(* IEC 61131-3 sources: deprecated-refusr-repo/GP/Main/samples (part 5) *)

(* ---- 3-MUX_sappy-ovals-yanks.st ---- *)
(*
This code implements a shuffled multiplexer with 3 control bits.
The control bits are: Data[2], Data[4], Data[1]
The input bits are: Data[6], Data[3], Data[5], Data[7], Data[9], Data[8], Data[10], Data[11]

The symbolic expression is:
(((((((~((~(D[2]) & ~(D[4])) & ~(D[1])) | D[6]) & (~((D[2] & ~(D[4])) & ~(D[1])) | D[3])) & (~((~(D[2]) & D[4]) & ~(D[1])) | D[5])) & (~((D[2] & D[4]) & ~(D[1])) | D[7])) & (~((~(D[2]) & ~(D[4])) & D[1]) | D[9])) & (~((D[2] & ~(D[4])) & D[1]) | D[8])) & (~((~(D[2]) & D[4]) & D[1]) | D[10])) & (~((D[2] & D[4]) & D[1]) | D[11])

*)

FUNCTION_BLOCK F_CollectInput
  VAR_IN_OUT
      Data : ARRAY[1..15] OF BOOL;
  END_VAR
  VAR_INPUT
      TICK  : BOOL := 0;
      IN1   : BOOL := 0;
      IN2   : BOOL := 0;
      IN3   : BOOL := 0;
      IN4   : BOOL := 0;
      IN5   : BOOL := 0;
      RESET : BOOL := FALSE;
  END_VAR
  VAR_OUTPUT
      Finished : BOOL;
  END_VAR
  VAR
      j    : USINT := 1;
      tock : BOOL  := 0;
  END_VAR
  IF NOT RESET AND tock = NOT TICK THEN
      Data[j]   := IN1;
      Data[j+1] := IN2;
      Data[j+2] := IN3;
      Data[j+3] := IN4;
      Data[j+4] := IN5;
      j := j + 5;
      tock := TICK;
  ELSE
      j := 1;
      tock := 0;
  END_IF;
  Finished := (j > 15);
END_FUNCTION_BLOCK

PROGRAM Boiler
  VAR
    Data  : ARRAY[1..15] OF BOOL;
    Ready : BOOL;
    CollectInput : F_CollectInput;
  END_VAR
  VAR
    TICK     AT %IX1.0 : BOOL;
    IN1      AT %IX0.3 : BOOL;
    IN2      AT %IX0.4 : BOOL;
    IN3      AT %IX0.5 : BOOL;
    IN4      AT %IX0.6 : BOOL;
    IN5      AT %IX0.7 : BOOL;
    OutReady AT %QX0.0 : BOOL := FALSE;
    FeedNext AT %QX0.1 : BOOL := FALSE;
    Out      AT %QX0.2 : BOOL;
  END_VAR
  CollectInput(TICK:=TICK, IN1:=IN1, IN2:=IN2, IN3:=IN3, IN4:=IN4, IN5:=IN5);
  Ready := CollectInput.Finished;
  FeedNext := 1;
  IF Ready THEN
    Out := (((((((((NOT (((NOT D[2]) AND (NOT D[4])) AND (NOT D[1]))) OR D[6]) AND ((NOT ((D[2] AND (NOT D[4])) AND (NOT D[1]))) OR D[3])) AND ((NOT (((NOT D[2]) AND D[4]) AND (NOT D[1]))) OR D[5])) AND ((NOT ((D[2] AND D[4]) AND (NOT D[1]))) OR D[7])) AND ((NOT (((NOT D[2]) AND (NOT D[4])) AND D[1])) OR D[9])) AND ((NOT ((D[2] AND (NOT D[4])) AND D[1])) OR D[8])) AND ((NOT (((NOT D[2]) AND D[4]) AND D[1])) OR D[10])) AND ((NOT ((D[2] AND D[4]) AND D[1])) OR D[11]));
    OutReady := 1;
    CollectInput(RESET:=TRUE);
  END_IF;
END_PROGRAM

CONFIGURATION Config0
  RESOURCE Res0 ON PLC
    TASK task0(INTERVAL := T#20ms,PRIORITY := 0);
    PROGRAM instance0 WITH task0 : Boiler;
  END_RESOURCE
END_CONFIGURATION

(* ---- 3-MUX_scale-wants-nifty.st ---- *)
(*
This code implements a shuffled multiplexer with 3 control bits.
The control bits are: Data[2], Data[3], Data[5]
The input bits are: Data[1], Data[8], Data[9], Data[7], Data[4], Data[10], Data[6], Data[11]

The symbolic expression is:
(((((((~((~(D[2]) & ~(D[3])) & ~(D[5])) | D[1]) & (~((D[2] & ~(D[3])) & ~(D[5])) | D[8])) & (~((~(D[2]) & D[3]) & ~(D[5])) | D[9])) & (~((D[2] & D[3]) & ~(D[5])) | D[7])) & (~((~(D[2]) & ~(D[3])) & D[5]) | D[4])) & (~((D[2] & ~(D[3])) & D[5]) | D[10])) & (~((~(D[2]) & D[3]) & D[5]) | D[6])) & (~((D[2] & D[3]) & D[5]) | D[11])

*)

FUNCTION_BLOCK F_CollectInput
  VAR_IN_OUT
      Data : ARRAY[1..15] OF BOOL;
  END_VAR
  VAR_INPUT
      TICK  : BOOL := 0;
      IN1   : BOOL := 0;
      IN2   : BOOL := 0;
      IN3   : BOOL := 0;
      IN4   : BOOL := 0;
      IN5   : BOOL := 0;
      RESET : BOOL := FALSE;
  END_VAR
  VAR_OUTPUT
      Finished : BOOL;
  END_VAR
  VAR
      j    : USINT := 1;
      tock : BOOL  := 0;
  END_VAR
  IF NOT RESET AND tock = NOT TICK THEN
      Data[j]   := IN1;
      Data[j+1] := IN2;
      Data[j+2] := IN3;
      Data[j+3] := IN4;
      Data[j+4] := IN5;
      j := j + 5;
      tock := TICK;
  ELSE
      j := 1;
      tock := 0;
  END_IF;
  Finished := (j > 15);
END_FUNCTION_BLOCK

PROGRAM Boiler
  VAR
    Data  : ARRAY[1..15] OF BOOL;
    Ready : BOOL;
    CollectInput : F_CollectInput;
  END_VAR
  VAR
    TICK     AT %IX1.0 : BOOL;
    IN1      AT %IX0.3 : BOOL;
    IN2      AT %IX0.4 : BOOL;
    IN3      AT %IX0.5 : BOOL;
    IN4      AT %IX0.6 : BOOL;
    IN5      AT %IX0.7 : BOOL;
    OutReady AT %QX0.0 : BOOL := FALSE;
    FeedNext AT %QX0.1 : BOOL := FALSE;
    Out      AT %QX0.2 : BOOL;
  END_VAR
  CollectInput(TICK:=TICK, IN1:=IN1, IN2:=IN2, IN3:=IN3, IN4:=IN4, IN5:=IN5);
  Ready := CollectInput.Finished;
  FeedNext := 1;
  IF Ready THEN
    Out := (((((((((NOT (((NOT D[2]) AND (NOT D[3])) AND (NOT D[5]))) OR D[1]) AND ((NOT ((D[2] AND (NOT D[3])) AND (NOT D[5]))) OR D[8])) AND ((NOT (((NOT D[2]) AND D[3]) AND (NOT D[5]))) OR D[9])) AND ((NOT ((D[2] AND D[3]) AND (NOT D[5]))) OR D[7])) AND ((NOT (((NOT D[2]) AND (NOT D[3])) AND D[5])) OR D[4])) AND ((NOT ((D[2] AND (NOT D[3])) AND D[5])) OR D[10])) AND ((NOT (((NOT D[2]) AND D[3]) AND D[5])) OR D[6])) AND ((NOT ((D[2] AND D[3]) AND D[5])) OR D[11]));
    OutReady := 1;
    CollectInput(RESET:=TRUE);
  END_IF;
END_PROGRAM

CONFIGURATION Config0
  RESOURCE Res0 ON PLC
    TASK task0(INTERVAL := T#20ms,PRIORITY := 0);
    PROGRAM instance0 WITH task0 : Boiler;
  END_RESOURCE
END_CONFIGURATION

(* ---- 3-MUX_scion-boxer-krona.st ---- *)
(*
This code implements a shuffled multiplexer with 3 control bits.
The control bits are: Data[3], Data[5], Data[4]
The input bits are: Data[1], Data[2], Data[9], Data[6], Data[10], Data[7], Data[11], Data[8]

The symbolic expression is:
(((((((~((~(D[3]) & ~(D[5])) & ~(D[4])) | D[1]) & (~((D[3] & ~(D[5])) & ~(D[4])) | D[2])) & (~((~(D[3]) & D[5]) & ~(D[4])) | D[9])) & (~((D[3] & D[5]) & ~(D[4])) | D[6])) & (~((~(D[3]) & ~(D[5])) & D[4]) | D[10])) & (~((D[3] & ~(D[5])) & D[4]) | D[7])) & (~((~(D[3]) & D[5]) & D[4]) | D[11])) & (~((D[3] & D[5]) & D[4]) | D[8])

*)

FUNCTION_BLOCK F_CollectInput
  VAR_IN_OUT
      Data : ARRAY[1..15] OF BOOL;
  END_VAR
  VAR_INPUT
      TICK  : BOOL := 0;
      IN1   : BOOL := 0;
      IN2   : BOOL := 0;
      IN3   : BOOL := 0;
      IN4   : BOOL := 0;
      IN5   : BOOL := 0;
      RESET : BOOL := FALSE;
  END_VAR
  VAR_OUTPUT
      Finished : BOOL;
  END_VAR
  VAR
      j    : USINT := 1;
      tock : BOOL  := 0;
  END_VAR
  IF NOT RESET AND tock = NOT TICK THEN
      Data[j]   := IN1;
      Data[j+1] := IN2;
      Data[j+2] := IN3;
      Data[j+3] := IN4;
      Data[j+4] := IN5;
      j := j + 5;
      tock := TICK;
  ELSE
      j := 1;
      tock := 0;
  END_IF;
  Finished := (j > 15);
END_FUNCTION_BLOCK

PROGRAM Boiler
  VAR
    Data  : ARRAY[1..15] OF BOOL;
    Ready : BOOL;
    CollectInput : F_CollectInput;
  END_VAR
  VAR
    TICK     AT %IX1.0 : BOOL;
    IN1      AT %IX0.3 : BOOL;
    IN2      AT %IX0.4 : BOOL;
    IN3      AT %IX0.5 : BOOL;
    IN4      AT %IX0.6 : BOOL;
    IN5      AT %IX0.7 : BOOL;
    OutReady AT %QX0.0 : BOOL := FALSE;
    FeedNext AT %QX0.1 : BOOL := FALSE;
    Out      AT %QX0.2 : BOOL;
  END_VAR
  CollectInput(TICK:=TICK, IN1:=IN1, IN2:=IN2, IN3:=IN3, IN4:=IN4, IN5:=IN5);
  Ready := CollectInput.Finished;
  FeedNext := 1;
  IF Ready THEN
    Out := (((((((((NOT (((NOT D[3]) AND (NOT D[5])) AND (NOT D[4]))) OR D[1]) AND ((NOT ((D[3] AND (NOT D[5])) AND (NOT D[4]))) OR D[2])) AND ((NOT (((NOT D[3]) AND D[5]) AND (NOT D[4]))) OR D[9])) AND ((NOT ((D[3] AND D[5]) AND (NOT D[4]))) OR D[6])) AND ((NOT (((NOT D[3]) AND (NOT D[5])) AND D[4])) OR D[10])) AND ((NOT ((D[3] AND (NOT D[5])) AND D[4])) OR D[7])) AND ((NOT (((NOT D[3]) AND D[5]) AND D[4])) OR D[11])) AND ((NOT ((D[3] AND D[5]) AND D[4])) OR D[8]));
    OutReady := 1;
    CollectInput(RESET:=TRUE);
  END_IF;
END_PROGRAM

CONFIGURATION Config0
  RESOURCE Res0 ON PLC
    TASK task0(INTERVAL := T#20ms,PRIORITY := 0);
    PROGRAM instance0 WITH task0 : Boiler;
  END_RESOURCE
END_CONFIGURATION

(* ---- 3-MUX_sects-chimp-tilth.st ---- *)
(*
This code implements a shuffled multiplexer with 3 control bits.
The control bits are: Data[2], Data[1], Data[5]
The input bits are: Data[3], Data[4], Data[6], Data[9], Data[7], Data[10], Data[11], Data[8]

The symbolic expression is:
(((((((~((~(D[2]) & ~(D[1])) & ~(D[5])) | D[3]) & (~((D[2] & ~(D[1])) & ~(D[5])) | D[4])) & (~((~(D[2]) & D[1]) & ~(D[5])) | D[6])) & (~((D[2] & D[1]) & ~(D[5])) | D[9])) & (~((~(D[2]) & ~(D[1])) & D[5]) | D[7])) & (~((D[2] & ~(D[1])) & D[5]) | D[10])) & (~((~(D[2]) & D[1]) & D[5]) | D[11])) & (~((D[2] & D[1]) & D[5]) | D[8])

*)

FUNCTION_BLOCK F_CollectInput
  VAR_IN_OUT
      Data : ARRAY[1..15] OF BOOL;
  END_VAR
  VAR_INPUT
      TICK  : BOOL := 0;
      IN1   : BOOL := 0;
      IN2   : BOOL := 0;
      IN3   : BOOL := 0;
      IN4   : BOOL := 0;
      IN5   : BOOL := 0;
      RESET : BOOL := FALSE;
  END_VAR
  VAR_OUTPUT
      Finished : BOOL;
  END_VAR
  VAR
      j    : USINT := 1;
      tock : BOOL  := 0;
  END_VAR
  IF NOT RESET AND tock = NOT TICK THEN
      Data[j]   := IN1;
      Data[j+1] := IN2;
      Data[j+2] := IN3;
      Data[j+3] := IN4;
      Data[j+4] := IN5;
      j := j + 5;
      tock := TICK;
  ELSE
      j := 1;
      tock := 0;
  END_IF;
  Finished := (j > 15);
END_FUNCTION_BLOCK

PROGRAM Boiler
  VAR
    Data  : ARRAY[1..15] OF BOOL;
    Ready : BOOL;
    CollectInput : F_CollectInput;
  END_VAR
  VAR
    TICK     AT %IX1.0 : BOOL;
    IN1      AT %IX0.3 : BOOL;
    IN2      AT %IX0.4 : BOOL;
    IN3      AT %IX0.5 : BOOL;
    IN4      AT %IX0.6 : BOOL;
    IN5      AT %IX0.7 : BOOL;
    OutReady AT %QX0.0 : BOOL := FALSE;
    FeedNext AT %QX0.1 : BOOL := FALSE;
    Out      AT %QX0.2 : BOOL;
  END_VAR
  CollectInput(TICK:=TICK, IN1:=IN1, IN2:=IN2, IN3:=IN3, IN4:=IN4, IN5:=IN5);
  Ready := CollectInput.Finished;
  FeedNext := 1;
  IF Ready THEN
    Out := (((((((((NOT (((NOT D[2]) AND (NOT D[1])) AND (NOT D[5]))) OR D[3]) AND ((NOT ((D[2] AND (NOT D[1])) AND (NOT D[5]))) OR D[4])) AND ((NOT (((NOT D[2]) AND D[1]) AND (NOT D[5]))) OR D[6])) AND ((NOT ((D[2] AND D[1]) AND (NOT D[5]))) OR D[9])) AND ((NOT (((NOT D[2]) AND (NOT D[1])) AND D[5])) OR D[7])) AND ((NOT ((D[2] AND (NOT D[1])) AND D[5])) OR D[10])) AND ((NOT (((NOT D[2]) AND D[1]) AND D[5])) OR D[11])) AND ((NOT ((D[2] AND D[1]) AND D[5])) OR D[8]));
    OutReady := 1;
    CollectInput(RESET:=TRUE);
  END_IF;
END_PROGRAM

CONFIGURATION Config0
  RESOURCE Res0 ON PLC
    TASK task0(INTERVAL := T#20ms,PRIORITY := 0);
    PROGRAM instance0 WITH task0 : Boiler;
  END_RESOURCE
END_CONFIGURATION

(* ---- 3-MUX_seems-zebra-casus.st ---- *)
(*
This code implements a shuffled multiplexer with 3 control bits.
The control bits are: Data[1], Data[2], Data[3]
The input bits are: Data[7], Data[5], Data[4], Data[6], Data[8], Data[9], Data[10], Data[11]

The symbolic expression is:
(((((((~((~(D[1]) & ~(D[2])) & ~(D[3])) | D[7]) & (~((D[1] & ~(D[2])) & ~(D[3])) | D[5])) & (~((~(D[1]) & D[2]) & ~(D[3])) | D[4])) & (~((D[1] & D[2]) & ~(D[3])) | D[6])) & (~((~(D[1]) & ~(D[2])) & D[3]) | D[8])) & (~((D[1] & ~(D[2])) & D[3]) | D[9])) & (~((~(D[1]) & D[2]) & D[3]) | D[10])) & (~((D[1] & D[2]) & D[3]) | D[11])

*)

FUNCTION_BLOCK F_CollectInput
  VAR_IN_OUT
      Data : ARRAY[1..15] OF BOOL;
  END_VAR
  VAR_INPUT
      TICK  : BOOL := 0;
      IN1   : BOOL := 0;
      IN2   : BOOL := 0;
      IN3   : BOOL := 0;
      IN4   : BOOL := 0;
      IN5   : BOOL := 0;
      RESET : BOOL := FALSE;
  END_VAR
  VAR_OUTPUT
      Finished : BOOL;
  END_VAR
  VAR
      j    : USINT := 1;
      tock : BOOL  := 0;
  END_VAR
  IF NOT RESET AND tock = NOT TICK THEN
      Data[j]   := IN1;
      Data[j+1] := IN2;
      Data[j+2] := IN3;
      Data[j+3] := IN4;
      Data[j+4] := IN5;
      j := j + 5;
      tock := TICK;
  ELSE
      j := 1;
      tock := 0;
  END_IF;
  Finished := (j > 15);
END_FUNCTION_BLOCK

PROGRAM Boiler
  VAR
    Data  : ARRAY[1..15] OF BOOL;
    Ready : BOOL;
    CollectInput : F_CollectInput;
  END_VAR
  VAR
    TICK     AT %IX1.0 : BOOL;
    IN1      AT %IX0.3 : BOOL;
    IN2      AT %IX0.4 : BOOL;
    IN3      AT %IX0.5 : BOOL;
    IN4      AT %IX0.6 : BOOL;
    IN5      AT %IX0.7 : BOOL;
    OutReady AT %QX0.0 : BOOL := FALSE;
    FeedNext AT %QX0.1 : BOOL := FALSE;
    Out      AT %QX0.2 : BOOL;
  END_VAR
  CollectInput(TICK:=TICK, IN1:=IN1, IN2:=IN2, IN3:=IN3, IN4:=IN4, IN5:=IN5);
  Ready := CollectInput.Finished;
  FeedNext := 1;
  IF Ready THEN
    Out := (((((((((NOT (((NOT D[1]) AND (NOT D[2])) AND (NOT D[3]))) OR D[7]) AND ((NOT ((D[1] AND (NOT D[2])) AND (NOT D[3]))) OR D[5])) AND ((NOT (((NOT D[1]) AND D[2]) AND (NOT D[3]))) OR D[4])) AND ((NOT ((D[1] AND D[2]) AND (NOT D[3]))) OR D[6])) AND ((NOT (((NOT D[1]) AND (NOT D[2])) AND D[3])) OR D[8])) AND ((NOT ((D[1] AND (NOT D[2])) AND D[3])) OR D[9])) AND ((NOT (((NOT D[1]) AND D[2]) AND D[3])) OR D[10])) AND ((NOT ((D[1] AND D[2]) AND D[3])) OR D[11]));
    OutReady := 1;
    CollectInput(RESET:=TRUE);
  END_IF;
END_PROGRAM

CONFIGURATION Config0
  RESOURCE Res0 ON PLC
    TASK task0(INTERVAL := T#20ms,PRIORITY := 0);
    PROGRAM instance0 WITH task0 : Boiler;
  END_RESOURCE
END_CONFIGURATION

(* ---- 3-MUX_shunt-caret-reedy.st ---- *)
(*
This code implements a shuffled multiplexer with 3 control bits.
The control bits are: Data[5], Data[3], Data[1]
The input bits are: Data[4], Data[6], Data[8], Data[7], Data[10], Data[11], Data[9], Data[2]

The symbolic expression is:
(((((((~((~(D[5]) & ~(D[3])) & ~(D[1])) | D[4]) & (~((D[5] & ~(D[3])) & ~(D[1])) | D[6])) & (~((~(D[5]) & D[3]) & ~(D[1])) | D[8])) & (~((D[5] & D[3]) & ~(D[1])) | D[7])) & (~((~(D[5]) & ~(D[3])) & D[1]) | D[10])) & (~((D[5] & ~(D[3])) & D[1]) | D[11])) & (~((~(D[5]) & D[3]) & D[1]) | D[9])) & (~((D[5] & D[3]) & D[1]) | D[2])

*)

FUNCTION_BLOCK F_CollectInput
  VAR_IN_OUT
      Data : ARRAY[1..15] OF BOOL;
  END_VAR
  VAR_INPUT
      TICK  : BOOL := 0;
      IN1   : BOOL := 0;
      IN2   : BOOL := 0;
      IN3   : BOOL := 0;
      IN4   : BOOL := 0;
      IN5   : BOOL := 0;
      RESET : BOOL := FALSE;
  END_VAR
  VAR_OUTPUT
      Finished : BOOL;
  END_VAR
  VAR
      j    : USINT := 1;
      tock : BOOL  := 0;
  END_VAR
  IF NOT RESET AND tock = NOT TICK THEN
      Data[j]   := IN1;
      Data[j+1] := IN2;
      Data[j+2] := IN3;
      Data[j+3] := IN4;
      Data[j+4] := IN5;
      j := j + 5;
      tock := TICK;
  ELSE
      j := 1;
      tock := 0;
  END_IF;
  Finished := (j > 15);
END_FUNCTION_BLOCK

PROGRAM Boiler
  VAR
    Data  : ARRAY[1..15] OF BOOL;
    Ready : BOOL;
    CollectInput : F_CollectInput;
  END_VAR
  VAR
    TICK     AT %IX1.0 : BOOL;
    IN1      AT %IX0.3 : BOOL;
    IN2      AT %IX0.4 : BOOL;
    IN3      AT %IX0.5 : BOOL;
    IN4      AT %IX0.6 : BOOL;
    IN5      AT %IX0.7 : BOOL;
    OutReady AT %QX0.0 : BOOL := FALSE;
    FeedNext AT %QX0.1 : BOOL := FALSE;
    Out      AT %QX0.2 : BOOL;
  END_VAR
  CollectInput(TICK:=TICK, IN1:=IN1, IN2:=IN2, IN3:=IN3, IN4:=IN4, IN5:=IN5);
  Ready := CollectInput.Finished;
  FeedNext := 1;
  IF Ready THEN
    Out := (((((((((NOT (((NOT D[5]) AND (NOT D[3])) AND (NOT D[1]))) OR D[4]) AND ((NOT ((D[5] AND (NOT D[3])) AND (NOT D[1]))) OR D[6])) AND ((NOT (((NOT D[5]) AND D[3]) AND (NOT D[1]))) OR D[8])) AND ((NOT ((D[5] AND D[3]) AND (NOT D[1]))) OR D[7])) AND ((NOT (((NOT D[5]) AND (NOT D[3])) AND D[1])) OR D[10])) AND ((NOT ((D[5] AND (NOT D[3])) AND D[1])) OR D[11])) AND ((NOT (((NOT D[5]) AND D[3]) AND D[1])) OR D[9])) AND ((NOT ((D[5] AND D[3]) AND D[1])) OR D[2]));
    OutReady := 1;
    CollectInput(RESET:=TRUE);
  END_IF;
END_PROGRAM

CONFIGURATION Config0
  RESOURCE Res0 ON PLC
    TASK task0(INTERVAL := T#20ms,PRIORITY := 0);
    PROGRAM instance0 WITH task0 : Boiler;
  END_RESOURCE
END_CONFIGURATION

(* ---- 3-MUX_slums-noted-letup.st ---- *)
(*
This code implements a shuffled multiplexer with 3 control bits.
The control bits are: Data[3], Data[4], Data[1]
The input bits are: Data[9], Data[2], Data[11], Data[5], Data[7], Data[8], Data[6], Data[10]

The symbolic expression is:
(((((((~((~(D[3]) & ~(D[4])) & ~(D[1])) | D[9]) & (~((D[3] & ~(D[4])) & ~(D[1])) | D[2])) & (~((~(D[3]) & D[4]) & ~(D[1])) | D[11])) & (~((D[3] & D[4]) & ~(D[1])) | D[5])) & (~((~(D[3]) & ~(D[4])) & D[1]) | D[7])) & (~((D[3] & ~(D[4])) & D[1]) | D[8])) & (~((~(D[3]) & D[4]) & D[1]) | D[6])) & (~((D[3] & D[4]) & D[1]) | D[10])

*)

FUNCTION_BLOCK F_CollectInput
  VAR_IN_OUT
      Data : ARRAY[1..15] OF BOOL;
  END_VAR
  VAR_INPUT
      TICK  : BOOL := 0;
      IN1   : BOOL := 0;
      IN2   : BOOL := 0;
      IN3   : BOOL := 0;
      IN4   : BOOL := 0;
      IN5   : BOOL := 0;
      RESET : BOOL := FALSE;
  END_VAR
  VAR_OUTPUT
      Finished : BOOL;
  END_VAR
  VAR
      j    : USINT := 1;
      tock : BOOL  := 0;
  END_VAR
  IF NOT RESET AND tock = NOT TICK THEN
      Data[j]   := IN1;
      Data[j+1] := IN2;
      Data[j+2] := IN3;
      Data[j+3] := IN4;
      Data[j+4] := IN5;
      j := j + 5;
      tock := TICK;
  ELSE
      j := 1;
      tock := 0;
  END_IF;
  Finished := (j > 15);
END_FUNCTION_BLOCK

PROGRAM Boiler
  VAR
    Data  : ARRAY[1..15] OF BOOL;
    Ready : BOOL;
    CollectInput : F_CollectInput;
  END_VAR
  VAR
    TICK     AT %IX1.0 : BOOL;
    IN1      AT %IX0.3 : BOOL;
    IN2      AT %IX0.4 : BOOL;
    IN3      AT %IX0.5 : BOOL;
    IN4      AT %IX0.6 : BOOL;
    IN5      AT %IX0.7 : BOOL;
    OutReady AT %QX0.0 : BOOL := FALSE;
    FeedNext AT %QX0.1 : BOOL := FALSE;
    Out      AT %QX0.2 : BOOL;
  END_VAR
  CollectInput(TICK:=TICK, IN1:=IN1, IN2:=IN2, IN3:=IN3, IN4:=IN4, IN5:=IN5);
  Ready := CollectInput.Finished;
  FeedNext := 1;
  IF Ready THEN
    Out := (((((((((NOT (((NOT D[3]) AND (NOT D[4])) AND (NOT D[1]))) OR D[9]) AND ((NOT ((D[3] AND (NOT D[4])) AND (NOT D[1]))) OR D[2])) AND ((NOT (((NOT D[3]) AND D[4]) AND (NOT D[1]))) OR D[11])) AND ((NOT ((D[3] AND D[4]) AND (NOT D[1]))) OR D[5])) AND ((NOT (((NOT D[3]) AND (NOT D[4])) AND D[1])) OR D[7])) AND ((NOT ((D[3] AND (NOT D[4])) AND D[1])) OR D[8])) AND ((NOT (((NOT D[3]) AND D[4]) AND D[1])) OR D[6])) AND ((NOT ((D[3] AND D[4]) AND D[1])) OR D[10]));
    OutReady := 1;
    CollectInput(RESET:=TRUE);
  END_IF;
END_PROGRAM

CONFIGURATION Config0
  RESOURCE Res0 ON PLC
    TASK task0(INTERVAL := T#20ms,PRIORITY := 0);
    PROGRAM instance0 WITH task0 : Boiler;
  END_RESOURCE
END_CONFIGURATION

(* ---- 3-MUX_sonny-vised-eying.st ---- *)
(*
This code implements a shuffled multiplexer with 3 control bits.
The control bits are: Data[2], Data[1], Data[4]
The input bits are: Data[3], Data[7], Data[6], Data[8], Data[5], Data[9], Data[11], Data[10]

The symbolic expression is:
(((((((~((~(D[2]) & ~(D[1])) & ~(D[4])) | D[3]) & (~((D[2] & ~(D[1])) & ~(D[4])) | D[7])) & (~((~(D[2]) & D[1]) & ~(D[4])) | D[6])) & (~((D[2] & D[1]) & ~(D[4])) | D[8])) & (~((~(D[2]) & ~(D[1])) & D[4]) | D[5])) & (~((D[2] & ~(D[1])) & D[4]) | D[9])) & (~((~(D[2]) & D[1]) & D[4]) | D[11])) & (~((D[2] & D[1]) & D[4]) | D[10])

*)

FUNCTION_BLOCK F_CollectInput
  VAR_IN_OUT
      Data : ARRAY[1..15] OF BOOL;
  END_VAR
  VAR_INPUT
      TICK  : BOOL := 0;
      IN1   : BOOL := 0;
      IN2   : BOOL := 0;
      IN3   : BOOL := 0;
      IN4   : BOOL := 0;
      IN5   : BOOL := 0;
      RESET : BOOL := FALSE;
  END_VAR
  VAR_OUTPUT
      Finished : BOOL;
  END_VAR
  VAR
      j    : USINT := 1;
      tock : BOOL  := 0;
  END_VAR
  IF NOT RESET AND tock = NOT TICK THEN
      Data[j]   := IN1;
      Data[j+1] := IN2;
      Data[j+2] := IN3;
      Data[j+3] := IN4;
      Data[j+4] := IN5;
      j := j + 5;
      tock := TICK;
  ELSE
      j := 1;
      tock := 0;
  END_IF;
  Finished := (j > 15);
END_FUNCTION_BLOCK

PROGRAM Boiler
  VAR
    Data  : ARRAY[1..15] OF BOOL;
    Ready : BOOL;
    CollectInput : F_CollectInput;
  END_VAR
  VAR
    TICK     AT %IX1.0 : BOOL;
    IN1      AT %IX0.3 : BOOL;
    IN2      AT %IX0.4 : BOOL;
    IN3      AT %IX0.5 : BOOL;
    IN4      AT %IX0.6 : BOOL;
    IN5      AT %IX0.7 : BOOL;
    OutReady AT %QX0.0 : BOOL := FALSE;
    FeedNext AT %QX0.1 : BOOL := FALSE;
    Out      AT %QX0.2 : BOOL;
  END_VAR
  CollectInput(TICK:=TICK, IN1:=IN1, IN2:=IN2, IN3:=IN3, IN4:=IN4, IN5:=IN5);
  Ready := CollectInput.Finished;
  FeedNext := 1;
  IF Ready THEN
    Out := (((((((((NOT (((NOT D[2]) AND (NOT D[1])) AND (NOT D[4]))) OR D[3]) AND ((NOT ((D[2] AND (NOT D[1])) AND (NOT D[4]))) OR D[7])) AND ((NOT (((NOT D[2]) AND D[1]) AND (NOT D[4]))) OR D[6])) AND ((NOT ((D[2] AND D[1]) AND (NOT D[4]))) OR D[8])) AND ((NOT (((NOT D[2]) AND (NOT D[1])) AND D[4])) OR D[5])) AND ((NOT ((D[2] AND (NOT D[1])) AND D[4])) OR D[9])) AND ((NOT (((NOT D[2]) AND D[1]) AND D[4])) OR D[11])) AND ((NOT ((D[2] AND D[1]) AND D[4])) OR D[10]));
    OutReady := 1;
    CollectInput(RESET:=TRUE);
  END_IF;
END_PROGRAM

CONFIGURATION Config0
  RESOURCE Res0 ON PLC
    TASK task0(INTERVAL := T#20ms,PRIORITY := 0);
    PROGRAM instance0 WITH task0 : Boiler;
  END_RESOURCE
END_CONFIGURATION

(* ---- 3-MUX_spark-lithe-swans.st ---- *)
(*
This code implements a shuffled multiplexer with 3 control bits.
The control bits are: Data[4], Data[3], Data[1]
The input bits are: Data[5], Data[6], Data[2], Data[7], Data[10], Data[8], Data[9], Data[11]

The symbolic expression is:
(((((((~((~(D[4]) & ~(D[3])) & ~(D[1])) | D[5]) & (~((D[4] & ~(D[3])) & ~(D[1])) | D[6])) & (~((~(D[4]) & D[3]) & ~(D[1])) | D[2])) & (~((D[4] & D[3]) & ~(D[1])) | D[7])) & (~((~(D[4]) & ~(D[3])) & D[1]) | D[10])) & (~((D[4] & ~(D[3])) & D[1]) | D[8])) & (~((~(D[4]) & D[3]) & D[1]) | D[9])) & (~((D[4] & D[3]) & D[1]) | D[11])

*)

FUNCTION_BLOCK F_CollectInput
  VAR_IN_OUT
      Data : ARRAY[1..15] OF BOOL;
  END_VAR
  VAR_INPUT
      TICK  : BOOL := 0;
      IN1   : BOOL := 0;
      IN2   : BOOL := 0;
      IN3   : BOOL := 0;
      IN4   : BOOL := 0;
      IN5   : BOOL := 0;
      RESET : BOOL := FALSE;
  END_VAR
  VAR_OUTPUT
      Finished : BOOL;
  END_VAR
  VAR
      j    : USINT := 1;
      tock : BOOL  := 0;
  END_VAR
  IF NOT RESET AND tock = NOT TICK THEN
      Data[j]   := IN1;
      Data[j+1] := IN2;
      Data[j+2] := IN3;
      Data[j+3] := IN4;
      Data[j+4] := IN5;
      j := j + 5;
      tock := TICK;
  ELSE
      j := 1;
      tock := 0;
  END_IF;
  Finished := (j > 15);
END_FUNCTION_BLOCK

PROGRAM Boiler
  VAR
    Data  : ARRAY[1..15] OF BOOL;
    Ready : BOOL;
    CollectInput : F_CollectInput;
  END_VAR
  VAR
    TICK     AT %IX1.0 : BOOL;
    IN1      AT %IX0.3 : BOOL;
    IN2      AT %IX0.4 : BOOL;
    IN3      AT %IX0.5 : BOOL;
    IN4      AT %IX0.6 : BOOL;
    IN5      AT %IX0.7 : BOOL;
    OutReady AT %QX0.0 : BOOL := FALSE;
    FeedNext AT %QX0.1 : BOOL := FALSE;
    Out      AT %QX0.2 : BOOL;
  END_VAR
  CollectInput(TICK:=TICK, IN1:=IN1, IN2:=IN2, IN3:=IN3, IN4:=IN4, IN5:=IN5);
  Ready := CollectInput.Finished;
  FeedNext := 1;
  IF Ready THEN
    Out := (((((((((NOT (((NOT D[4]) AND (NOT D[3])) AND (NOT D[1]))) OR D[5]) AND ((NOT ((D[4] AND (NOT D[3])) AND (NOT D[1]))) OR D[6])) AND ((NOT (((NOT D[4]) AND D[3]) AND (NOT D[1]))) OR D[2])) AND ((NOT ((D[4] AND D[3]) AND (NOT D[1]))) OR D[7])) AND ((NOT (((NOT D[4]) AND (NOT D[3])) AND D[1])) OR D[10])) AND ((NOT ((D[4] AND (NOT D[3])) AND D[1])) OR D[8])) AND ((NOT (((NOT D[4]) AND D[3]) AND D[1])) OR D[9])) AND ((NOT ((D[4] AND D[3]) AND D[1])) OR D[11]));
    OutReady := 1;
    CollectInput(RESET:=TRUE);
  END_IF;
END_PROGRAM

CONFIGURATION Config0
  RESOURCE Res0 ON PLC
    TASK task0(INTERVAL := T#20ms,PRIORITY := 0);
    PROGRAM instance0 WITH task0 : Boiler;
  END_RESOURCE
END_CONFIGURATION

(* ---- 3-MUX_spoof-lawns-sylph.st ---- *)
(*
This code implements a shuffled multiplexer with 3 control bits.
The control bits are: Data[2], Data[1], Data[3]
The input bits are: Data[4], Data[7], Data[8], Data[5], Data[9], Data[6], Data[10], Data[11]

The symbolic expression is:
(((((((~((~(D[2]) & ~(D[1])) & ~(D[3])) | D[4]) & (~((D[2] & ~(D[1])) & ~(D[3])) | D[7])) & (~((~(D[2]) & D[1]) & ~(D[3])) | D[8])) & (~((D[2] & D[1]) & ~(D[3])) | D[5])) & (~((~(D[2]) & ~(D[1])) & D[3]) | D[9])) & (~((D[2] & ~(D[1])) & D[3]) | D[6])) & (~((~(D[2]) & D[1]) & D[3]) | D[10])) & (~((D[2] & D[1]) & D[3]) | D[11])

*)

FUNCTION_BLOCK F_CollectInput
  VAR_IN_OUT
      Data : ARRAY[1..15] OF BOOL;
  END_VAR
  VAR_INPUT
      TICK  : BOOL := 0;
      IN1   : BOOL := 0;
      IN2   : BOOL := 0;
      IN3   : BOOL := 0;
      IN4   : BOOL := 0;
      IN5   : BOOL := 0;
      RESET : BOOL := FALSE;
  END_VAR
  VAR_OUTPUT
      Finished : BOOL;
  END_VAR
  VAR
      j    : USINT := 1;
      tock : BOOL  := 0;
  END_VAR
  IF NOT RESET AND tock = NOT TICK THEN
      Data[j]   := IN1;
      Data[j+1] := IN2;
      Data[j+2] := IN3;
      Data[j+3] := IN4;
      Data[j+4] := IN5;
      j := j + 5;
      tock := TICK;
  ELSE
      j := 1;
      tock := 0;
  END_IF;
  Finished := (j > 15);
END_FUNCTION_BLOCK

PROGRAM Boiler
  VAR
    Data  : ARRAY[1..15] OF BOOL;
    Ready : BOOL;
    CollectInput : F_CollectInput;
  END_VAR
  VAR
    TICK     AT %IX1.0 : BOOL;
    IN1      AT %IX0.3 : BOOL;
    IN2      AT %IX0.4 : BOOL;
    IN3      AT %IX0.5 : BOOL;
    IN4      AT %IX0.6 : BOOL;
    IN5      AT %IX0.7 : BOOL;
    OutReady AT %QX0.0 : BOOL := FALSE;
    FeedNext AT %QX0.1 : BOOL := FALSE;
    Out      AT %QX0.2 : BOOL;
  END_VAR
  CollectInput(TICK:=TICK, IN1:=IN1, IN2:=IN2, IN3:=IN3, IN4:=IN4, IN5:=IN5);
  Ready := CollectInput.Finished;
  FeedNext := 1;
  IF Ready THEN
    Out := (((((((((NOT (((NOT D[2]) AND (NOT D[1])) AND (NOT D[3]))) OR D[4]) AND ((NOT ((D[2] AND (NOT D[1])) AND (NOT D[3]))) OR D[7])) AND ((NOT (((NOT D[2]) AND D[1]) AND (NOT D[3]))) OR D[8])) AND ((NOT ((D[2] AND D[1]) AND (NOT D[3]))) OR D[5])) AND ((NOT (((NOT D[2]) AND (NOT D[1])) AND D[3])) OR D[9])) AND ((NOT ((D[2] AND (NOT D[1])) AND D[3])) OR D[6])) AND ((NOT (((NOT D[2]) AND D[1]) AND D[3])) OR D[10])) AND ((NOT ((D[2] AND D[1]) AND D[3])) OR D[11]));
    OutReady := 1;
    CollectInput(RESET:=TRUE);
  END_IF;
END_PROGRAM

CONFIGURATION Config0
  RESOURCE Res0 ON PLC
    TASK task0(INTERVAL := T#20ms,PRIORITY := 0);
    PROGRAM instance0 WITH task0 : Boiler;
  END_RESOURCE
END_CONFIGURATION

(* ---- 3-MUX_steer-patsy-bored.st ---- *)
(*
This code implements a shuffled multiplexer with 3 control bits.
The control bits are: Data[3], Data[1], Data[2]
The input bits are: Data[5], Data[4], Data[6], Data[9], Data[7], Data[11], Data[8], Data[10]

The symbolic expression is:
(((((((~((~(D[3]) & ~(D[1])) & ~(D[2])) | D[5]) & (~((D[3] & ~(D[1])) & ~(D[2])) | D[4])) & (~((~(D[3]) & D[1]) & ~(D[2])) | D[6])) & (~((D[3] & D[1]) & ~(D[2])) | D[9])) & (~((~(D[3]) & ~(D[1])) & D[2]) | D[7])) & (~((D[3] & ~(D[1])) & D[2]) | D[11])) & (~((~(D[3]) & D[1]) & D[2]) | D[8])) & (~((D[3] & D[1]) & D[2]) | D[10])

*)

FUNCTION_BLOCK F_CollectInput
  VAR_IN_OUT
      Data : ARRAY[1..15] OF BOOL;
  END_VAR
  VAR_INPUT
      TICK  : BOOL := 0;
      IN1   : BOOL := 0;
      IN2   : BOOL := 0;
      IN3   : BOOL := 0;
      IN4   : BOOL := 0;
      IN5   : BOOL := 0;
      RESET : BOOL := FALSE;
  END_VAR
  VAR_OUTPUT
      Finished : BOOL;
  END_VAR
  VAR
      j    : USINT := 1;
      tock : BOOL  := 0;
  END_VAR
  IF NOT RESET AND tock = NOT TICK THEN
      Data[j]   := IN1;
      Data[j+1] := IN2;
      Data[j+2] := IN3;
      Data[j+3] := IN4;
      Data[j+4] := IN5;
      j := j + 5;
      tock := TICK;
  ELSE
      j := 1;
      tock := 0;
  END_IF;
  Finished := (j > 15);
END_FUNCTION_BLOCK

PROGRAM Boiler
  VAR
    Data  : ARRAY[1..15] OF BOOL;
    Ready : BOOL;
    CollectInput : F_CollectInput;
  END_VAR
  VAR
    TICK     AT %IX1.0 : BOOL;
    IN1      AT %IX0.3 : BOOL;
    IN2      AT %IX0.4 : BOOL;
    IN3      AT %IX0.5 : BOOL;
    IN4      AT %IX0.6 : BOOL;
    IN5      AT %IX0.7 : BOOL;
    OutReady AT %QX0.0 : BOOL := FALSE;
    FeedNext AT %QX0.1 : BOOL := FALSE;
    Out      AT %QX0.2 : BOOL;
  END_VAR
  CollectInput(TICK:=TICK, IN1:=IN1, IN2:=IN2, IN3:=IN3, IN4:=IN4, IN5:=IN5);
  Ready := CollectInput.Finished;
  FeedNext := 1;
  IF Ready THEN
    Out := (((((((((NOT (((NOT D[3]) AND (NOT D[1])) AND (NOT D[2]))) OR D[5]) AND ((NOT ((D[3] AND (NOT D[1])) AND (NOT D[2]))) OR D[4])) AND ((NOT (((NOT D[3]) AND D[1]) AND (NOT D[2]))) OR D[6])) AND ((NOT ((D[3] AND D[1]) AND (NOT D[2]))) OR D[9])) AND ((NOT (((NOT D[3]) AND (NOT D[1])) AND D[2])) OR D[7])) AND ((NOT ((D[3] AND (NOT D[1])) AND D[2])) OR D[11])) AND ((NOT (((NOT D[3]) AND D[1]) AND D[2])) OR D[8])) AND ((NOT ((D[3] AND D[1]) AND D[2])) OR D[10]));
    OutReady := 1;
    CollectInput(RESET:=TRUE);
  END_IF;
END_PROGRAM

CONFIGURATION Config0
  RESOURCE Res0 ON PLC
    TASK task0(INTERVAL := T#20ms,PRIORITY := 0);
    PROGRAM instance0 WITH task0 : Boiler;
  END_RESOURCE
END_CONFIGURATION

(* ---- 3-MUX_sting-scurf-goons.st ---- *)
(*
This code implements a shuffled multiplexer with 3 control bits.
The control bits are: Data[1], Data[3], Data[2]
The input bits are: Data[4], Data[6], Data[5], Data[8], Data[7], Data[9], Data[10], Data[11]

The symbolic expression is:
(((((((~((~(D[1]) & ~(D[3])) & ~(D[2])) | D[4]) & (~((D[1] & ~(D[3])) & ~(D[2])) | D[6])) & (~((~(D[1]) & D[3]) & ~(D[2])) | D[5])) & (~((D[1] & D[3]) & ~(D[2])) | D[8])) & (~((~(D[1]) & ~(D[3])) & D[2]) | D[7])) & (~((D[1] & ~(D[3])) & D[2]) | D[9])) & (~((~(D[1]) & D[3]) & D[2]) | D[10])) & (~((D[1] & D[3]) & D[2]) | D[11])

*)

FUNCTION_BLOCK F_CollectInput
  VAR_IN_OUT
      Data : ARRAY[1..15] OF BOOL;
  END_VAR
  VAR_INPUT
      TICK  : BOOL := 0;
      IN1   : BOOL := 0;
      IN2   : BOOL := 0;
      IN3   : BOOL := 0;
      IN4   : BOOL := 0;
      IN5   : BOOL := 0;
      RESET : BOOL := FALSE;
  END_VAR
  VAR_OUTPUT
      Finished : BOOL;
  END_VAR
  VAR
      j    : USINT := 1;
      tock : BOOL  := 0;
  END_VAR
  IF NOT RESET AND tock = NOT TICK THEN
      Data[j]   := IN1;
      Data[j+1] := IN2;
      Data[j+2] := IN3;
      Data[j+3] := IN4;
      Data[j+4] := IN5;
      j := j + 5;
      tock := TICK;
  ELSE
      j := 1;
      tock := 0;
  END_IF;
  Finished := (j > 15);
END_FUNCTION_BLOCK

PROGRAM Boiler
  VAR
    Data  : ARRAY[1..15] OF BOOL;
    Ready : BOOL;
    CollectInput : F_CollectInput;
  END_VAR
  VAR
    TICK     AT %IX1.0 : BOOL;
    IN1      AT %IX0.3 : BOOL;
    IN2      AT %IX0.4 : BOOL;
    IN3      AT %IX0.5 : BOOL;
    IN4      AT %IX0.6 : BOOL;
    IN5      AT %IX0.7 : BOOL;
    OutReady AT %QX0.0 : BOOL := FALSE;
    FeedNext AT %QX0.1 : BOOL := FALSE;
    Out      AT %QX0.2 : BOOL;
  END_VAR
  CollectInput(TICK:=TICK, IN1:=IN1, IN2:=IN2, IN3:=IN3, IN4:=IN4, IN5:=IN5);
  Ready := CollectInput.Finished;
  FeedNext := 1;
  IF Ready THEN
    Out := (((((((((NOT (((NOT D[1]) AND (NOT D[3])) AND (NOT D[2]))) OR D[4]) AND ((NOT ((D[1] AND (NOT D[3])) AND (NOT D[2]))) OR D[6])) AND ((NOT (((NOT D[1]) AND D[3]) AND (NOT D[2]))) OR D[5])) AND ((NOT ((D[1] AND D[3]) AND (NOT D[2]))) OR D[8])) AND ((NOT (((NOT D[1]) AND (NOT D[3])) AND D[2])) OR D[7])) AND ((NOT ((D[1] AND (NOT D[3])) AND D[2])) OR D[9])) AND ((NOT (((NOT D[1]) AND D[3]) AND D[2])) OR D[10])) AND ((NOT ((D[1] AND D[3]) AND D[2])) OR D[11]));
    OutReady := 1;
    CollectInput(RESET:=TRUE);
  END_IF;
END_PROGRAM

CONFIGURATION Config0
  RESOURCE Res0 ON PLC
    TASK task0(INTERVAL := T#20ms,PRIORITY := 0);
    PROGRAM instance0 WITH task0 : Boiler;
  END_RESOURCE
END_CONFIGURATION

(* ---- 3-MUX_stoop-pubis-sitar.st ---- *)
(*
This code implements a shuffled multiplexer with 3 control bits.
The control bits are: Data[1], Data[2], Data[4]
The input bits are: Data[6], Data[3], Data[5], Data[9], Data[8], Data[7], Data[11], Data[10]

The symbolic expression is:
(((((((~((~(D[1]) & ~(D[2])) & ~(D[4])) | D[6]) & (~((D[1] & ~(D[2])) & ~(D[4])) | D[3])) & (~((~(D[1]) & D[2]) & ~(D[4])) | D[5])) & (~((D[1] & D[2]) & ~(D[4])) | D[9])) & (~((~(D[1]) & ~(D[2])) & D[4]) | D[8])) & (~((D[1] & ~(D[2])) & D[4]) | D[7])) & (~((~(D[1]) & D[2]) & D[4]) | D[11])) & (~((D[1] & D[2]) & D[4]) | D[10])

*)

FUNCTION_BLOCK F_CollectInput
  VAR_IN_OUT
      Data : ARRAY[1..15] OF BOOL;
  END_VAR
  VAR_INPUT
      TICK  : BOOL := 0;
      IN1   : BOOL := 0;
      IN2   : BOOL := 0;
      IN3   : BOOL := 0;
      IN4   : BOOL := 0;
      IN5   : BOOL := 0;
      RESET : BOOL := FALSE;
  END_VAR
  VAR_OUTPUT
      Finished : BOOL;
  END_VAR
  VAR
      j    : USINT := 1;
      tock : BOOL  := 0;
  END_VAR
  IF NOT RESET AND tock = NOT TICK THEN
      Data[j]   := IN1;
      Data[j+1] := IN2;
      Data[j+2] := IN3;
      Data[j+3] := IN4;
      Data[j+4] := IN5;
      j := j + 5;
      tock := TICK;
  ELSE
      j := 1;
      tock := 0;
  END_IF;
  Finished := (j > 15);
END_FUNCTION_BLOCK

PROGRAM Boiler
  VAR
    Data  : ARRAY[1..15] OF BOOL;
    Ready : BOOL;
    CollectInput : F_CollectInput;
  END_VAR
  VAR
    TICK     AT %IX1.0 : BOOL;
    IN1      AT %IX0.3 : BOOL;
    IN2      AT %IX0.4 : BOOL;
    IN3      AT %IX0.5 : BOOL;
    IN4      AT %IX0.6 : BOOL;
    IN5      AT %IX0.7 : BOOL;
    OutReady AT %QX0.0 : BOOL := FALSE;
    FeedNext AT %QX0.1 : BOOL := FALSE;
    Out      AT %QX0.2 : BOOL;
  END_VAR
  CollectInput(TICK:=TICK, IN1:=IN1, IN2:=IN2, IN3:=IN3, IN4:=IN4, IN5:=IN5);
  Ready := CollectInput.Finished;
  FeedNext := 1;
  IF Ready THEN
    Out := (((((((((NOT (((NOT D[1]) AND (NOT D[2])) AND (NOT D[4]))) OR D[6]) AND ((NOT ((D[1] AND (NOT D[2])) AND (NOT D[4]))) OR D[3])) AND ((NOT (((NOT D[1]) AND D[2]) AND (NOT D[4]))) OR D[5])) AND ((NOT ((D[1] AND D[2]) AND (NOT D[4]))) OR D[9])) AND ((NOT (((NOT D[1]) AND (NOT D[2])) AND D[4])) OR D[8])) AND ((NOT ((D[1] AND (NOT D[2])) AND D[4])) OR D[7])) AND ((NOT (((NOT D[1]) AND D[2]) AND D[4])) OR D[11])) AND ((NOT ((D[1] AND D[2]) AND D[4])) OR D[10]));
    OutReady := 1;
    CollectInput(RESET:=TRUE);
  END_IF;
END_PROGRAM

CONFIGURATION Config0
  RESOURCE Res0 ON PLC
    TASK task0(INTERVAL := T#20ms,PRIORITY := 0);
    PROGRAM instance0 WITH task0 : Boiler;
  END_RESOURCE
END_CONFIGURATION

(* ---- 3-MUX_swart-fulls-comic.st ---- *)
(*
This code implements a shuffled multiplexer with 3 control bits.
The control bits are: Data[3], Data[1], Data[4]
The input bits are: Data[2], Data[5], Data[6], Data[8], Data[7], Data[11], Data[10], Data[9]

The symbolic expression is:
(((((((~((~(D[3]) & ~(D[1])) & ~(D[4])) | D[2]) & (~((D[3] & ~(D[1])) & ~(D[4])) | D[5])) & (~((~(D[3]) & D[1]) & ~(D[4])) | D[6])) & (~((D[3] & D[1]) & ~(D[4])) | D[8])) & (~((~(D[3]) & ~(D[1])) & D[4]) | D[7])) & (~((D[3] & ~(D[1])) & D[4]) | D[11])) & (~((~(D[3]) & D[1]) & D[4]) | D[10])) & (~((D[3] & D[1]) & D[4]) | D[9])

*)

FUNCTION_BLOCK F_CollectInput
  VAR_IN_OUT
      Data : ARRAY[1..15] OF BOOL;
  END_VAR
  VAR_INPUT
      TICK  : BOOL := 0;
      IN1   : BOOL := 0;
      IN2   : BOOL := 0;
      IN3   : BOOL := 0;
      IN4   : BOOL := 0;
      IN5   : BOOL := 0;
      RESET : BOOL := FALSE;
  END_VAR
  VAR_OUTPUT
      Finished : BOOL;
  END_VAR
  VAR
      j    : USINT := 1;
      tock : BOOL  := 0;
  END_VAR
  IF NOT RESET AND tock = NOT TICK THEN
      Data[j]   := IN1;
      Data[j+1] := IN2;
      Data[j+2] := IN3;
      Data[j+3] := IN4;
      Data[j+4] := IN5;
      j := j + 5;
      tock := TICK;
  ELSE
      j := 1;
      tock := 0;
  END_IF;
  Finished := (j > 15);
END_FUNCTION_BLOCK

PROGRAM Boiler
  VAR
    Data  : ARRAY[1..15] OF BOOL;
    Ready : BOOL;
    CollectInput : F_CollectInput;
  END_VAR
  VAR
    TICK     AT %IX1.0 : BOOL;
    IN1      AT %IX0.3 : BOOL;
    IN2      AT %IX0.4 : BOOL;
    IN3      AT %IX0.5 : BOOL;
    IN4      AT %IX0.6 : BOOL;
    IN5      AT %IX0.7 : BOOL;
    OutReady AT %QX0.0 : BOOL := FALSE;
    FeedNext AT %QX0.1 : BOOL := FALSE;
    Out      AT %QX0.2 : BOOL;
  END_VAR
  CollectInput(TICK:=TICK, IN1:=IN1, IN2:=IN2, IN3:=IN3, IN4:=IN4, IN5:=IN5);
  Ready := CollectInput.Finished;
  FeedNext := 1;
  IF Ready THEN
    Out := (((((((((NOT (((NOT D[3]) AND (NOT D[1])) AND (NOT D[4]))) OR D[2]) AND ((NOT ((D[3] AND (NOT D[1])) AND (NOT D[4]))) OR D[5])) AND ((NOT (((NOT D[3]) AND D[1]) AND (NOT D[4]))) OR D[6])) AND ((NOT ((D[3] AND D[1]) AND (NOT D[4]))) OR D[8])) AND ((NOT (((NOT D[3]) AND (NOT D[1])) AND D[4])) OR D[7])) AND ((NOT ((D[3] AND (NOT D[1])) AND D[4])) OR D[11])) AND ((NOT (((NOT D[3]) AND D[1]) AND D[4])) OR D[10])) AND ((NOT ((D[3] AND D[1]) AND D[4])) OR D[9]));
    OutReady := 1;
    CollectInput(RESET:=TRUE);
  END_IF;
END_PROGRAM

CONFIGURATION Config0
  RESOURCE Res0 ON PLC
    TASK task0(INTERVAL := T#20ms,PRIORITY := 0);
    PROGRAM instance0 WITH task0 : Boiler;
  END_RESOURCE
END_CONFIGURATION

(* ---- 3-MUX_terce-henge-chino.st ---- *)
(*
This code implements a shuffled multiplexer with 3 control bits.
The control bits are: Data[3], Data[4], Data[5]
The input bits are: Data[2], Data[6], Data[7], Data[1], Data[8], Data[11], Data[10], Data[9]

The symbolic expression is:
(((((((~((~(D[3]) & ~(D[4])) & ~(D[5])) | D[2]) & (~((D[3] & ~(D[4])) & ~(D[5])) | D[6])) & (~((~(D[3]) & D[4]) & ~(D[5])) | D[7])) & (~((D[3] & D[4]) & ~(D[5])) | D[1])) & (~((~(D[3]) & ~(D[4])) & D[5]) | D[8])) & (~((D[3] & ~(D[4])) & D[5]) | D[11])) & (~((~(D[3]) & D[4]) & D[5]) | D[10])) & (~((D[3] & D[4]) & D[5]) | D[9])

*)

FUNCTION_BLOCK F_CollectInput
  VAR_IN_OUT
      Data : ARRAY[1..15] OF BOOL;
  END_VAR
  VAR_INPUT
      TICK  : BOOL := 0;
      IN1   : BOOL := 0;
      IN2   : BOOL := 0;
      IN3   : BOOL := 0;
      IN4   : BOOL := 0;
      IN5   : BOOL := 0;
      RESET : BOOL := FALSE;
  END_VAR
  VAR_OUTPUT
      Finished : BOOL;
  END_VAR
  VAR
      j    : USINT := 1;
      tock : BOOL  := 0;
  END_VAR
  IF NOT RESET AND tock = NOT TICK THEN
      Data[j]   := IN1;
      Data[j+1] := IN2;
      Data[j+2] := IN3;
      Data[j+3] := IN4;
      Data[j+4] := IN5;
      j := j + 5;
      tock := TICK;
  ELSE
      j := 1;
      tock := 0;
  END_IF;
  Finished := (j > 15);
END_FUNCTION_BLOCK

PROGRAM Boiler
  VAR
    Data  : ARRAY[1..15] OF BOOL;
    Ready : BOOL;
    CollectInput : F_CollectInput;
  END_VAR
  VAR
    TICK     AT %IX1.0 : BOOL;
    IN1      AT %IX0.3 : BOOL;
    IN2      AT %IX0.4 : BOOL;
    IN3      AT %IX0.5 : BOOL;
    IN4      AT %IX0.6 : BOOL;
    IN5      AT %IX0.7 : BOOL;
    OutReady AT %QX0.0 : BOOL := FALSE;
    FeedNext AT %QX0.1 : BOOL := FALSE;
    Out      AT %QX0.2 : BOOL;
  END_VAR
  CollectInput(TICK:=TICK, IN1:=IN1, IN2:=IN2, IN3:=IN3, IN4:=IN4, IN5:=IN5);
  Ready := CollectInput.Finished;
  FeedNext := 1;
  IF Ready THEN
    Out := (((((((((NOT (((NOT D[3]) AND (NOT D[4])) AND (NOT D[5]))) OR D[2]) AND ((NOT ((D[3] AND (NOT D[4])) AND (NOT D[5]))) OR D[6])) AND ((NOT (((NOT D[3]) AND D[4]) AND (NOT D[5]))) OR D[7])) AND ((NOT ((D[3] AND D[4]) AND (NOT D[5]))) OR D[1])) AND ((NOT (((NOT D[3]) AND (NOT D[4])) AND D[5])) OR D[8])) AND ((NOT ((D[3] AND (NOT D[4])) AND D[5])) OR D[11])) AND ((NOT (((NOT D[3]) AND D[4]) AND D[5])) OR D[10])) AND ((NOT ((D[3] AND D[4]) AND D[5])) OR D[9]));
    OutReady := 1;
    CollectInput(RESET:=TRUE);
  END_IF;
END_PROGRAM

CONFIGURATION Config0
  RESOURCE Res0 ON PLC
    TASK task0(INTERVAL := T#20ms,PRIORITY := 0);
    PROGRAM instance0 WITH task0 : Boiler;
  END_RESOURCE
END_CONFIGURATION

(* ---- 3-MUX_thank-chums-segue.st ---- *)
(*
This code implements a shuffled multiplexer with 3 control bits.
The control bits are: Data[1], Data[3], Data[4]
The input bits are: Data[5], Data[2], Data[7], Data[6], Data[9], Data[8], Data[11], Data[10]

The symbolic expression is:
(((((((~((~(D[1]) & ~(D[3])) & ~(D[4])) | D[5]) & (~((D[1] & ~(D[3])) & ~(D[4])) | D[2])) & (~((~(D[1]) & D[3]) & ~(D[4])) | D[7])) & (~((D[1] & D[3]) & ~(D[4])) | D[6])) & (~((~(D[1]) & ~(D[3])) & D[4]) | D[9])) & (~((D[1] & ~(D[3])) & D[4]) | D[8])) & (~((~(D[1]) & D[3]) & D[4]) | D[11])) & (~((D[1] & D[3]) & D[4]) | D[10])

*)

FUNCTION_BLOCK F_CollectInput
  VAR_IN_OUT
      Data : ARRAY[1..15] OF BOOL;
  END_VAR
  VAR_INPUT
      TICK  : BOOL := 0;
      IN1   : BOOL := 0;
      IN2   : BOOL := 0;
      IN3   : BOOL := 0;
      IN4   : BOOL := 0;
      IN5   : BOOL := 0;
      RESET : BOOL := FALSE;
  END_VAR
  VAR_OUTPUT
      Finished : BOOL;
  END_VAR
  VAR
      j    : USINT := 1;
      tock : BOOL  := 0;
  END_VAR
  IF NOT RESET AND tock = NOT TICK THEN
      Data[j]   := IN1;
      Data[j+1] := IN2;
      Data[j+2] := IN3;
      Data[j+3] := IN4;
      Data[j+4] := IN5;
      j := j + 5;
      tock := TICK;
  ELSE
      j := 1;
      tock := 0;
  END_IF;
  Finished := (j > 15);
END_FUNCTION_BLOCK

PROGRAM Boiler
  VAR
    Data  : ARRAY[1..15] OF BOOL;
    Ready : BOOL;
    CollectInput : F_CollectInput;
  END_VAR
  VAR
    TICK     AT %IX1.0 : BOOL;
    IN1      AT %IX0.3 : BOOL;
    IN2      AT %IX0.4 : BOOL;
    IN3      AT %IX0.5 : BOOL;
    IN4      AT %IX0.6 : BOOL;
    IN5      AT %IX0.7 : BOOL;
    OutReady AT %QX0.0 : BOOL := FALSE;
    FeedNext AT %QX0.1 : BOOL := FALSE;
    Out      AT %QX0.2 : BOOL;
  END_VAR
  CollectInput(TICK:=TICK, IN1:=IN1, IN2:=IN2, IN3:=IN3, IN4:=IN4, IN5:=IN5);
  Ready := CollectInput.Finished;
  FeedNext := 1;
  IF Ready THEN
    Out := (((((((((NOT (((NOT D[1]) AND (NOT D[3])) AND (NOT D[4]))) OR D[5]) AND ((NOT ((D[1] AND (NOT D[3])) AND (NOT D[4]))) OR D[2])) AND ((NOT (((NOT D[1]) AND D[3]) AND (NOT D[4]))) OR D[7])) AND ((NOT ((D[1] AND D[3]) AND (NOT D[4]))) OR D[6])) AND ((NOT (((NOT D[1]) AND (NOT D[3])) AND D[4])) OR D[9])) AND ((NOT ((D[1] AND (NOT D[3])) AND D[4])) OR D[8])) AND ((NOT (((NOT D[1]) AND D[3]) AND D[4])) OR D[11])) AND ((NOT ((D[1] AND D[3]) AND D[4])) OR D[10]));
    OutReady := 1;
    CollectInput(RESET:=TRUE);
  END_IF;
END_PROGRAM

CONFIGURATION Config0
  RESOURCE Res0 ON PLC
    TASK task0(INTERVAL := T#20ms,PRIORITY := 0);
    PROGRAM instance0 WITH task0 : Boiler;
  END_RESOURCE
END_CONFIGURATION

(* ---- 3-MUX_throw-salve-gears.st ---- *)
(*
This code implements a shuffled multiplexer with 3 control bits.
The control bits are: Data[1], Data[4], Data[2]
The input bits are: Data[8], Data[10], Data[3], Data[7], Data[5], Data[9], Data[6], Data[11]

The symbolic expression is:
(((((((~((~(D[1]) & ~(D[4])) & ~(D[2])) | D[8]) & (~((D[1] & ~(D[4])) & ~(D[2])) | D[10])) & (~((~(D[1]) & D[4]) & ~(D[2])) | D[3])) & (~((D[1] & D[4]) & ~(D[2])) | D[7])) & (~((~(D[1]) & ~(D[4])) & D[2]) | D[5])) & (~((D[1] & ~(D[4])) & D[2]) | D[9])) & (~((~(D[1]) & D[4]) & D[2]) | D[6])) & (~((D[1] & D[4]) & D[2]) | D[11])

*)

FUNCTION_BLOCK F_CollectInput
  VAR_IN_OUT
      Data : ARRAY[1..15] OF BOOL;
  END_VAR
  VAR_INPUT
      TICK  : BOOL := 0;
      IN1   : BOOL := 0;
      IN2   : BOOL := 0;
      IN3   : BOOL := 0;
      IN4   : BOOL := 0;
      IN5   : BOOL := 0;
      RESET : BOOL := FALSE;
  END_VAR
  VAR_OUTPUT
      Finished : BOOL;
  END_VAR
  VAR
      j    : USINT := 1;
      tock : BOOL  := 0;
  END_VAR
  IF NOT RESET AND tock = NOT TICK THEN
      Data[j]   := IN1;
      Data[j+1] := IN2;
      Data[j+2] := IN3;
      Data[j+3] := IN4;
      Data[j+4] := IN5;
      j := j + 5;
      tock := TICK;
  ELSE
      j := 1;
      tock := 0;
  END_IF;
  Finished := (j > 15);
END_FUNCTION_BLOCK

PROGRAM Boiler
  VAR
    Data  : ARRAY[1..15] OF BOOL;
    Ready : BOOL;
    CollectInput : F_CollectInput;
  END_VAR
  VAR
    TICK     AT %IX1.0 : BOOL;
    IN1      AT %IX0.3 : BOOL;
    IN2      AT %IX0.4 : BOOL;
    IN3      AT %IX0.5 : BOOL;
    IN4      AT %IX0.6 : BOOL;
    IN5      AT %IX0.7 : BOOL;
    OutReady AT %QX0.0 : BOOL := FALSE;
    FeedNext AT %QX0.1 : BOOL := FALSE;
    Out      AT %QX0.2 : BOOL;
  END_VAR
  CollectInput(TICK:=TICK, IN1:=IN1, IN2:=IN2, IN3:=IN3, IN4:=IN4, IN5:=IN5);
  Ready := CollectInput.Finished;
  FeedNext := 1;
  IF Ready THEN
    Out := (((((((((NOT (((NOT D[1]) AND (NOT D[4])) AND (NOT D[2]))) OR D[8]) AND ((NOT ((D[1] AND (NOT D[4])) AND (NOT D[2]))) OR D[10])) AND ((NOT (((NOT D[1]) AND D[4]) AND (NOT D[2]))) OR D[3])) AND ((NOT ((D[1] AND D[4]) AND (NOT D[2]))) OR D[7])) AND ((NOT (((NOT D[1]) AND (NOT D[4])) AND D[2])) OR D[5])) AND ((NOT ((D[1] AND (NOT D[4])) AND D[2])) OR D[9])) AND ((NOT (((NOT D[1]) AND D[4]) AND D[2])) OR D[6])) AND ((NOT ((D[1] AND D[4]) AND D[2])) OR D[11]));
    OutReady := 1;
    CollectInput(RESET:=TRUE);
  END_IF;
END_PROGRAM

CONFIGURATION Config0
  RESOURCE Res0 ON PLC
    TASK task0(INTERVAL := T#20ms,PRIORITY := 0);
    PROGRAM instance0 WITH task0 : Boiler;
  END_RESOURCE
END_CONFIGURATION

(* ---- 3-MUX_torus-nudes-psalm.st ---- *)
(*
This code implements a shuffled multiplexer with 3 control bits.
The control bits are: Data[4], Data[2], Data[1]
The input bits are: Data[3], Data[5], Data[8], Data[6], Data[11], Data[7], Data[9], Data[10]

The symbolic expression is:
(((((((~((~(D[4]) & ~(D[2])) & ~(D[1])) | D[3]) & (~((D[4] & ~(D[2])) & ~(D[1])) | D[5])) & (~((~(D[4]) & D[2]) & ~(D[1])) | D[8])) & (~((D[4] & D[2]) & ~(D[1])) | D[6])) & (~((~(D[4]) & ~(D[2])) & D[1]) | D[11])) & (~((D[4] & ~(D[2])) & D[1]) | D[7])) & (~((~(D[4]) & D[2]) & D[1]) | D[9])) & (~((D[4] & D[2]) & D[1]) | D[10])

*)

FUNCTION_BLOCK F_CollectInput
  VAR_IN_OUT
      Data : ARRAY[1..15] OF BOOL;
  END_VAR
  VAR_INPUT
      TICK  : BOOL := 0;
      IN1   : BOOL := 0;
      IN2   : BOOL := 0;
      IN3   : BOOL := 0;
      IN4   : BOOL := 0;
      IN5   : BOOL := 0;
      RESET : BOOL := FALSE;
  END_VAR
  VAR_OUTPUT
      Finished : BOOL;
  END_VAR
  VAR
      j    : USINT := 1;
      tock : BOOL  := 0;
  END_VAR
  IF NOT RESET AND tock = NOT TICK THEN
      Data[j]   := IN1;
      Data[j+1] := IN2;
      Data[j+2] := IN3;
      Data[j+3] := IN4;
      Data[j+4] := IN5;
      j := j + 5;
      tock := TICK;
  ELSE
      j := 1;
      tock := 0;
  END_IF;
  Finished := (j > 15);
END_FUNCTION_BLOCK

PROGRAM Boiler
  VAR
    Data  : ARRAY[1..15] OF BOOL;
    Ready : BOOL;
    CollectInput : F_CollectInput;
  END_VAR
  VAR
    TICK     AT %IX1.0 : BOOL;
    IN1      AT %IX0.3 : BOOL;
    IN2      AT %IX0.4 : BOOL;
    IN3      AT %IX0.5 : BOOL;
    IN4      AT %IX0.6 : BOOL;
    IN5      AT %IX0.7 : BOOL;
    OutReady AT %QX0.0 : BOOL := FALSE;
    FeedNext AT %QX0.1 : BOOL := FALSE;
    Out      AT %QX0.2 : BOOL;
  END_VAR
  CollectInput(TICK:=TICK, IN1:=IN1, IN2:=IN2, IN3:=IN3, IN4:=IN4, IN5:=IN5);
  Ready := CollectInput.Finished;
  FeedNext := 1;
  IF Ready THEN
    Out := (((((((((NOT (((NOT D[4]) AND (NOT D[2])) AND (NOT D[1]))) OR D[3]) AND ((NOT ((D[4] AND (NOT D[2])) AND (NOT D[1]))) OR D[5])) AND ((NOT (((NOT D[4]) AND D[2]) AND (NOT D[1]))) OR D[8])) AND ((NOT ((D[4] AND D[2]) AND (NOT D[1]))) OR D[6])) AND ((NOT (((NOT D[4]) AND (NOT D[2])) AND D[1])) OR D[11])) AND ((NOT ((D[4] AND (NOT D[2])) AND D[1])) OR D[7])) AND ((NOT (((NOT D[4]) AND D[2]) AND D[1])) OR D[9])) AND ((NOT ((D[4] AND D[2]) AND D[1])) OR D[10]));
    OutReady := 1;
    CollectInput(RESET:=TRUE);
  END_IF;
END_PROGRAM

CONFIGURATION Config0
  RESOURCE Res0 ON PLC
    TASK task0(INTERVAL := T#20ms,PRIORITY := 0);
    PROGRAM instance0 WITH task0 : Boiler;
  END_RESOURCE
END_CONFIGURATION

(* ---- 3-MUX_trees-ruddy-caped.st ---- *)
(*
This code implements a shuffled multiplexer with 3 control bits.
The control bits are: Data[5], Data[1], Data[2]
The input bits are: Data[9], Data[6], Data[3], Data[4], Data[7], Data[8], Data[10], Data[11]

The symbolic expression is:
(((((((~((~(D[5]) & ~(D[1])) & ~(D[2])) | D[9]) & (~((D[5] & ~(D[1])) & ~(D[2])) | D[6])) & (~((~(D[5]) & D[1]) & ~(D[2])) | D[3])) & (~((D[5] & D[1]) & ~(D[2])) | D[4])) & (~((~(D[5]) & ~(D[1])) & D[2]) | D[7])) & (~((D[5] & ~(D[1])) & D[2]) | D[8])) & (~((~(D[5]) & D[1]) & D[2]) | D[10])) & (~((D[5] & D[1]) & D[2]) | D[11])

*)

FUNCTION_BLOCK F_CollectInput
  VAR_IN_OUT
      Data : ARRAY[1..15] OF BOOL;
  END_VAR
  VAR_INPUT
      TICK  : BOOL := 0;
      IN1   : BOOL := 0;
      IN2   : BOOL := 0;
      IN3   : BOOL := 0;
      IN4   : BOOL := 0;
      IN5   : BOOL := 0;
      RESET : BOOL := FALSE;
  END_VAR
  VAR_OUTPUT
      Finished : BOOL;
  END_VAR
  VAR
      j    : USINT := 1;
      tock : BOOL  := 0;
  END_VAR
  IF NOT RESET AND tock = NOT TICK THEN
      Data[j]   := IN1;
      Data[j+1] := IN2;
      Data[j+2] := IN3;
      Data[j+3] := IN4;
      Data[j+4] := IN5;
      j := j + 5;
      tock := TICK;
  ELSE
      j := 1;
      tock := 0;
  END_IF;
  Finished := (j > 15);
END_FUNCTION_BLOCK

PROGRAM Boiler
  VAR
    Data  : ARRAY[1..15] OF BOOL;
    Ready : BOOL;
    CollectInput : F_CollectInput;
  END_VAR
  VAR
    TICK     AT %IX1.0 : BOOL;
    IN1      AT %IX0.3 : BOOL;
    IN2      AT %IX0.4 : BOOL;
    IN3      AT %IX0.5 : BOOL;
    IN4      AT %IX0.6 : BOOL;
    IN5      AT %IX0.7 : BOOL;
    OutReady AT %QX0.0 : BOOL := FALSE;
    FeedNext AT %QX0.1 : BOOL := FALSE;
    Out      AT %QX0.2 : BOOL;
  END_VAR
  CollectInput(TICK:=TICK, IN1:=IN1, IN2:=IN2, IN3:=IN3, IN4:=IN4, IN5:=IN5);
  Ready := CollectInput.Finished;
  FeedNext := 1;
  IF Ready THEN
    Out := (((((((((NOT (((NOT D[5]) AND (NOT D[1])) AND (NOT D[2]))) OR D[9]) AND ((NOT ((D[5] AND (NOT D[1])) AND (NOT D[2]))) OR D[6])) AND ((NOT (((NOT D[5]) AND D[1]) AND (NOT D[2]))) OR D[3])) AND ((NOT ((D[5] AND D[1]) AND (NOT D[2]))) OR D[4])) AND ((NOT (((NOT D[5]) AND (NOT D[1])) AND D[2])) OR D[7])) AND ((NOT ((D[5] AND (NOT D[1])) AND D[2])) OR D[8])) AND ((NOT (((NOT D[5]) AND D[1]) AND D[2])) OR D[10])) AND ((NOT ((D[5] AND D[1]) AND D[2])) OR D[11]));
    OutReady := 1;
    CollectInput(RESET:=TRUE);
  END_IF;
END_PROGRAM

CONFIGURATION Config0
  RESOURCE Res0 ON PLC
    TASK task0(INTERVAL := T#20ms,PRIORITY := 0);
    PROGRAM instance0 WITH task0 : Boiler;
  END_RESOURCE
END_CONFIGURATION

(* ---- 3-MUX_tumor-abbot-jokes.st ---- *)
(*
This code implements a shuffled multiplexer with 3 control bits.
The control bits are: Data[3], Data[1], Data[2]
The input bits are: Data[4], Data[5], Data[10], Data[6], Data[7], Data[11], Data[9], Data[8]

The symbolic expression is:
(((((((~((~(D[3]) & ~(D[1])) & ~(D[2])) | D[4]) & (~((D[3] & ~(D[1])) & ~(D[2])) | D[5])) & (~((~(D[3]) & D[1]) & ~(D[2])) | D[10])) & (~((D[3] & D[1]) & ~(D[2])) | D[6])) & (~((~(D[3]) & ~(D[1])) & D[2]) | D[7])) & (~((D[3] & ~(D[1])) & D[2]) | D[11])) & (~((~(D[3]) & D[1]) & D[2]) | D[9])) & (~((D[3] & D[1]) & D[2]) | D[8])

*)

FUNCTION_BLOCK F_CollectInput
  VAR_IN_OUT
      Data : ARRAY[1..15] OF BOOL;
  END_VAR
  VAR_INPUT
      TICK  : BOOL := 0;
      IN1   : BOOL := 0;
      IN2   : BOOL := 0;
      IN3   : BOOL := 0;
      IN4   : BOOL := 0;
      IN5   : BOOL := 0;
      RESET : BOOL := FALSE;
  END_VAR
  VAR_OUTPUT
      Finished : BOOL;
  END_VAR
  VAR
      j    : USINT := 1;
      tock : BOOL  := 0;
  END_VAR
  IF NOT RESET AND tock = NOT TICK THEN
      Data[j]   := IN1;
      Data[j+1] := IN2;
      Data[j+2] := IN3;
      Data[j+3] := IN4;
      Data[j+4] := IN5;
      j := j + 5;
      tock := TICK;
  ELSE
      j := 1;
      tock := 0;
  END_IF;
  Finished := (j > 15);
END_FUNCTION_BLOCK

PROGRAM Boiler
  VAR
    Data  : ARRAY[1..15] OF BOOL;
    Ready : BOOL;
    CollectInput : F_CollectInput;
  END_VAR
  VAR
    TICK     AT %IX1.0 : BOOL;
    IN1      AT %IX0.3 : BOOL;
    IN2      AT %IX0.4 : BOOL;
    IN3      AT %IX0.5 : BOOL;
    IN4      AT %IX0.6 : BOOL;
    IN5      AT %IX0.7 : BOOL;
    OutReady AT %QX0.0 : BOOL := FALSE;
    FeedNext AT %QX0.1 : BOOL := FALSE;
    Out      AT %QX0.2 : BOOL;
  END_VAR
  CollectInput(TICK:=TICK, IN1:=IN1, IN2:=IN2, IN3:=IN3, IN4:=IN4, IN5:=IN5);
  Ready := CollectInput.Finished;
  FeedNext := 1;
  IF Ready THEN
    Out := (((((((((NOT (((NOT D[3]) AND (NOT D[1])) AND (NOT D[2]))) OR D[4]) AND ((NOT ((D[3] AND (NOT D[1])) AND (NOT D[2]))) OR D[5])) AND ((NOT (((NOT D[3]) AND D[1]) AND (NOT D[2]))) OR D[10])) AND ((NOT ((D[3] AND D[1]) AND (NOT D[2]))) OR D[6])) AND ((NOT (((NOT D[3]) AND (NOT D[1])) AND D[2])) OR D[7])) AND ((NOT ((D[3] AND (NOT D[1])) AND D[2])) OR D[11])) AND ((NOT (((NOT D[3]) AND D[1]) AND D[2])) OR D[9])) AND ((NOT ((D[3] AND D[1]) AND D[2])) OR D[8]));
    OutReady := 1;
    CollectInput(RESET:=TRUE);
  END_IF;
END_PROGRAM

CONFIGURATION Config0
  RESOURCE Res0 ON PLC
    TASK task0(INTERVAL := T#20ms,PRIORITY := 0);
    PROGRAM instance0 WITH task0 : Boiler;
  END_RESOURCE
END_CONFIGURATION

(* ---- 3-MUX_twink-spoil-comic.st ---- *)
(*
This code implements a shuffled multiplexer with 3 control bits.
The control bits are: Data[4], Data[3], Data[2]
The input bits are: Data[7], Data[1], Data[8], Data[9], Data[10], Data[5], Data[11], Data[6]

The symbolic expression is:
(((((((~((~(D[4]) & ~(D[3])) & ~(D[2])) | D[7]) & (~((D[4] & ~(D[3])) & ~(D[2])) | D[1])) & (~((~(D[4]) & D[3]) & ~(D[2])) | D[8])) & (~((D[4] & D[3]) & ~(D[2])) | D[9])) & (~((~(D[4]) & ~(D[3])) & D[2]) | D[10])) & (~((D[4] & ~(D[3])) & D[2]) | D[5])) & (~((~(D[4]) & D[3]) & D[2]) | D[11])) & (~((D[4] & D[3]) & D[2]) | D[6])

*)

FUNCTION_BLOCK F_CollectInput
  VAR_IN_OUT
      Data : ARRAY[1..15] OF BOOL;
  END_VAR
  VAR_INPUT
      TICK  : BOOL := 0;
      IN1   : BOOL := 0;
      IN2   : BOOL := 0;
      IN3   : BOOL := 0;
      IN4   : BOOL := 0;
      IN5   : BOOL := 0;
      RESET : BOOL := FALSE;
  END_VAR
  VAR_OUTPUT
      Finished : BOOL;
  END_VAR
  VAR
      j    : USINT := 1;
      tock : BOOL  := 0;
  END_VAR
  IF NOT RESET AND tock = NOT TICK THEN
      Data[j]   := IN1;
      Data[j+1] := IN2;
      Data[j+2] := IN3;
      Data[j+3] := IN4;
      Data[j+4] := IN5;
      j := j + 5;
      tock := TICK;
  ELSE
      j := 1;
      tock := 0;
  END_IF;
  Finished := (j > 15);
END_FUNCTION_BLOCK

PROGRAM Boiler
  VAR
    Data  : ARRAY[1..15] OF BOOL;
    Ready : BOOL;
    CollectInput : F_CollectInput;
  END_VAR
  VAR
    TICK     AT %IX1.0 : BOOL;
    IN1      AT %IX0.3 : BOOL;
    IN2      AT %IX0.4 : BOOL;
    IN3      AT %IX0.5 : BOOL;
    IN4      AT %IX0.6 : BOOL;
    IN5      AT %IX0.7 : BOOL;
    OutReady AT %QX0.0 : BOOL := FALSE;
    FeedNext AT %QX0.1 : BOOL := FALSE;
    Out      AT %QX0.2 : BOOL;
  END_VAR
  CollectInput(TICK:=TICK, IN1:=IN1, IN2:=IN2, IN3:=IN3, IN4:=IN4, IN5:=IN5);
  Ready := CollectInput.Finished;
  FeedNext := 1;
  IF Ready THEN
    Out := (((((((((NOT (((NOT D[4]) AND (NOT D[3])) AND (NOT D[2]))) OR D[7]) AND ((NOT ((D[4] AND (NOT D[3])) AND (NOT D[2]))) OR D[1])) AND ((NOT (((NOT D[4]) AND D[3]) AND (NOT D[2]))) OR D[8])) AND ((NOT ((D[4] AND D[3]) AND (NOT D[2]))) OR D[9])) AND ((NOT (((NOT D[4]) AND (NOT D[3])) AND D[2])) OR D[10])) AND ((NOT ((D[4] AND (NOT D[3])) AND D[2])) OR D[5])) AND ((NOT (((NOT D[4]) AND D[3]) AND D[2])) OR D[11])) AND ((NOT ((D[4] AND D[3]) AND D[2])) OR D[6]));
    OutReady := 1;
    CollectInput(RESET:=TRUE);
  END_IF;
END_PROGRAM

CONFIGURATION Config0
  RESOURCE Res0 ON PLC
    TASK task0(INTERVAL := T#20ms,PRIORITY := 0);
    PROGRAM instance0 WITH task0 : Boiler;
  END_RESOURCE
END_CONFIGURATION

(* ---- 3-MUX_ultra-arson-aport.st ---- *)
(*
This code implements a shuffled multiplexer with 3 control bits.
The control bits are: Data[2], Data[1], Data[9]
The input bits are: Data[3], Data[7], Data[8], Data[6], Data[4], Data[5], Data[11], Data[10]

The symbolic expression is:
(((((((~((~(D[2]) & ~(D[1])) & ~(D[9])) | D[3]) & (~((D[2] & ~(D[1])) & ~(D[9])) | D[7])) & (~((~(D[2]) & D[1]) & ~(D[9])) | D[8])) & (~((D[2] & D[1]) & ~(D[9])) | D[6])) & (~((~(D[2]) & ~(D[1])) & D[9]) | D[4])) & (~((D[2] & ~(D[1])) & D[9]) | D[5])) & (~((~(D[2]) & D[1]) & D[9]) | D[11])) & (~((D[2] & D[1]) & D[9]) | D[10])

*)

FUNCTION_BLOCK F_CollectInput
  VAR_IN_OUT
      Data : ARRAY[1..15] OF BOOL;
  END_VAR
  VAR_INPUT
      TICK  : BOOL := 0;
      IN1   : BOOL := 0;
      IN2   : BOOL := 0;
      IN3   : BOOL := 0;
      IN4   : BOOL := 0;
      IN5   : BOOL := 0;
      RESET : BOOL := FALSE;
  END_VAR
  VAR_OUTPUT
      Finished : BOOL;
  END_VAR
  VAR
      j    : USINT := 1;
      tock : BOOL  := 0;
  END_VAR
  IF NOT RESET AND tock = NOT TICK THEN
      Data[j]   := IN1;
      Data[j+1] := IN2;
      Data[j+2] := IN3;
      Data[j+3] := IN4;
      Data[j+4] := IN5;
      j := j + 5;
      tock := TICK;
  ELSE
      j := 1;
      tock := 0;
  END_IF;
  Finished := (j > 15);
END_FUNCTION_BLOCK

PROGRAM Boiler
  VAR
    Data  : ARRAY[1..15] OF BOOL;
    Ready : BOOL;
    CollectInput : F_CollectInput;
  END_VAR
  VAR
    TICK     AT %IX1.0 : BOOL;
    IN1      AT %IX0.3 : BOOL;
    IN2      AT %IX0.4 : BOOL;
    IN3      AT %IX0.5 : BOOL;
    IN4      AT %IX0.6 : BOOL;
    IN5      AT %IX0.7 : BOOL;
    OutReady AT %QX0.0 : BOOL := FALSE;
    FeedNext AT %QX0.1 : BOOL := FALSE;
    Out      AT %QX0.2 : BOOL;
  END_VAR
  CollectInput(TICK:=TICK, IN1:=IN1, IN2:=IN2, IN3:=IN3, IN4:=IN4, IN5:=IN5);
  Ready := CollectInput.Finished;
  FeedNext := 1;
  IF Ready THEN
    Out := (((((((((NOT (((NOT D[2]) AND (NOT D[1])) AND (NOT D[9]))) OR D[3]) AND ((NOT ((D[2] AND (NOT D[1])) AND (NOT D[9]))) OR D[7])) AND ((NOT (((NOT D[2]) AND D[1]) AND (NOT D[9]))) OR D[8])) AND ((NOT ((D[2] AND D[1]) AND (NOT D[9]))) OR D[6])) AND ((NOT (((NOT D[2]) AND (NOT D[1])) AND D[9])) OR D[4])) AND ((NOT ((D[2] AND (NOT D[1])) AND D[9])) OR D[5])) AND ((NOT (((NOT D[2]) AND D[1]) AND D[9])) OR D[11])) AND ((NOT ((D[2] AND D[1]) AND D[9])) OR D[10]));
    OutReady := 1;
    CollectInput(RESET:=TRUE);
  END_IF;
END_PROGRAM

CONFIGURATION Config0
  RESOURCE Res0 ON PLC
    TASK task0(INTERVAL := T#20ms,PRIORITY := 0);
    PROGRAM instance0 WITH task0 : Boiler;
  END_RESOURCE
END_CONFIGURATION

(* ---- 3-MUX_unjam-gauge-honks.st ---- *)
(*
This code implements a shuffled multiplexer with 3 control bits.
The control bits are: Data[7], Data[2], Data[3]
The input bits are: Data[1], Data[5], Data[4], Data[8], Data[9], Data[11], Data[6], Data[10]

The symbolic expression is:
(((((((~((~(D[7]) & ~(D[2])) & ~(D[3])) | D[1]) & (~((D[7] & ~(D[2])) & ~(D[3])) | D[5])) & (~((~(D[7]) & D[2]) & ~(D[3])) | D[4])) & (~((D[7] & D[2]) & ~(D[3])) | D[8])) & (~((~(D[7]) & ~(D[2])) & D[3]) | D[9])) & (~((D[7] & ~(D[2])) & D[3]) | D[11])) & (~((~(D[7]) & D[2]) & D[3]) | D[6])) & (~((D[7] & D[2]) & D[3]) | D[10])

*)

FUNCTION_BLOCK F_CollectInput
  VAR_IN_OUT
      Data : ARRAY[1..15] OF BOOL;
  END_VAR
  VAR_INPUT
      TICK  : BOOL := 0;
      IN1   : BOOL := 0;
      IN2   : BOOL := 0;
      IN3   : BOOL := 0;
      IN4   : BOOL := 0;
      IN5   : BOOL := 0;
      RESET : BOOL := FALSE;
  END_VAR
  VAR_OUTPUT
      Finished : BOOL;
  END_VAR
  VAR
      j    : USINT := 1;
      tock : BOOL  := 0;
  END_VAR
  IF NOT RESET AND tock = NOT TICK THEN
      Data[j]   := IN1;
      Data[j+1] := IN2;
      Data[j+2] := IN3;
      Data[j+3] := IN4;
      Data[j+4] := IN5;
      j := j + 5;
      tock := TICK;
  ELSE
      j := 1;
      tock := 0;
  END_IF;
  Finished := (j > 15);
END_FUNCTION_BLOCK

PROGRAM Boiler
  VAR
    Data  : ARRAY[1..15] OF BOOL;
    Ready : BOOL;
    CollectInput : F_CollectInput;
  END_VAR
  VAR
    TICK     AT %IX1.0 : BOOL;
    IN1      AT %IX0.3 : BOOL;
    IN2      AT %IX0.4 : BOOL;
    IN3      AT %IX0.5 : BOOL;
    IN4      AT %IX0.6 : BOOL;
    IN5      AT %IX0.7 : BOOL;
    OutReady AT %QX0.0 : BOOL := FALSE;
    FeedNext AT %QX0.1 : BOOL := FALSE;
    Out      AT %QX0.2 : BOOL;
  END_VAR
  CollectInput(TICK:=TICK, IN1:=IN1, IN2:=IN2, IN3:=IN3, IN4:=IN4, IN5:=IN5);
  Ready := CollectInput.Finished;
  FeedNext := 1;
  IF Ready THEN
    Out := (((((((((NOT (((NOT D[7]) AND (NOT D[2])) AND (NOT D[3]))) OR D[1]) AND ((NOT ((D[7] AND (NOT D[2])) AND (NOT D[3]))) OR D[5])) AND ((NOT (((NOT D[7]) AND D[2]) AND (NOT D[3]))) OR D[4])) AND ((NOT ((D[7] AND D[2]) AND (NOT D[3]))) OR D[8])) AND ((NOT (((NOT D[7]) AND (NOT D[2])) AND D[3])) OR D[9])) AND ((NOT ((D[7] AND (NOT D[2])) AND D[3])) OR D[11])) AND ((NOT (((NOT D[7]) AND D[2]) AND D[3])) OR D[6])) AND ((NOT ((D[7] AND D[2]) AND D[3])) OR D[10]));
    OutReady := 1;
    CollectInput(RESET:=TRUE);
  END_IF;
END_PROGRAM

CONFIGURATION Config0
  RESOURCE Res0 ON PLC
    TASK task0(INTERVAL := T#20ms,PRIORITY := 0);
    PROGRAM instance0 WITH task0 : Boiler;
  END_RESOURCE
END_CONFIGURATION

(* ---- 3-MUX_unlit-talcs-halts.st ---- *)
(*
This code implements a shuffled multiplexer with 3 control bits.
The control bits are: Data[1], Data[2], Data[3]
The input bits are: Data[4], Data[5], Data[6], Data[7], Data[8], Data[10], Data[9], Data[11]

The symbolic expression is:
(((((((~((~(D[1]) & ~(D[2])) & ~(D[3])) | D[4]) & (~((D[1] & ~(D[2])) & ~(D[3])) | D[5])) & (~((~(D[1]) & D[2]) & ~(D[3])) | D[6])) & (~((D[1] & D[2]) & ~(D[3])) | D[7])) & (~((~(D[1]) & ~(D[2])) & D[3]) | D[8])) & (~((D[1] & ~(D[2])) & D[3]) | D[10])) & (~((~(D[1]) & D[2]) & D[3]) | D[9])) & (~((D[1] & D[2]) & D[3]) | D[11])

*)

FUNCTION_BLOCK F_CollectInput
  VAR_IN_OUT
      Data : ARRAY[1..15] OF BOOL;
  END_VAR
  VAR_INPUT
      TICK  : BOOL := 0;
      IN1   : BOOL := 0;
      IN2   : BOOL := 0;
      IN3   : BOOL := 0;
      IN4   : BOOL := 0;
      IN5   : BOOL := 0;
      RESET : BOOL := FALSE;
  END_VAR
  VAR_OUTPUT
      Finished : BOOL;
  END_VAR
  VAR
      j    : USINT := 1;
      tock : BOOL  := 0;
  END_VAR
  IF NOT RESET AND tock = NOT TICK THEN
      Data[j]   := IN1;
      Data[j+1] := IN2;
      Data[j+2] := IN3;
      Data[j+3] := IN4;
      Data[j+4] := IN5;
      j := j + 5;
      tock := TICK;
  ELSE
      j := 1;
      tock := 0;
  END_IF;
  Finished := (j > 15);
END_FUNCTION_BLOCK

PROGRAM Boiler
  VAR
    Data  : ARRAY[1..15] OF BOOL;
    Ready : BOOL;
    CollectInput : F_CollectInput;
  END_VAR
  VAR
    TICK     AT %IX1.0 : BOOL;
    IN1      AT %IX0.3 : BOOL;
    IN2      AT %IX0.4 : BOOL;
    IN3      AT %IX0.5 : BOOL;
    IN4      AT %IX0.6 : BOOL;
    IN5      AT %IX0.7 : BOOL;
    OutReady AT %QX0.0 : BOOL := FALSE;
    FeedNext AT %QX0.1 : BOOL := FALSE;
    Out      AT %QX0.2 : BOOL;
  END_VAR
  CollectInput(TICK:=TICK, IN1:=IN1, IN2:=IN2, IN3:=IN3, IN4:=IN4, IN5:=IN5);
  Ready := CollectInput.Finished;
  FeedNext := 1;
  IF Ready THEN
    Out := (((((((((NOT (((NOT D[1]) AND (NOT D[2])) AND (NOT D[3]))) OR D[4]) AND ((NOT ((D[1] AND (NOT D[2])) AND (NOT D[3]))) OR D[5])) AND ((NOT (((NOT D[1]) AND D[2]) AND (NOT D[3]))) OR D[6])) AND ((NOT ((D[1] AND D[2]) AND (NOT D[3]))) OR D[7])) AND ((NOT (((NOT D[1]) AND (NOT D[2])) AND D[3])) OR D[8])) AND ((NOT ((D[1] AND (NOT D[2])) AND D[3])) OR D[10])) AND ((NOT (((NOT D[1]) AND D[2]) AND D[3])) OR D[9])) AND ((NOT ((D[1] AND D[2]) AND D[3])) OR D[11]));
    OutReady := 1;
    CollectInput(RESET:=TRUE);
  END_IF;
END_PROGRAM

CONFIGURATION Config0
  RESOURCE Res0 ON PLC
    TASK task0(INTERVAL := T#20ms,PRIORITY := 0);
    PROGRAM instance0 WITH task0 : Boiler;
  END_RESOURCE
END_CONFIGURATION

(* ---- 3-MUX_usury-mooch-duets.st ---- *)
(*
This code implements a shuffled multiplexer with 3 control bits.
The control bits are: Data[2], Data[1], Data[4]
The input bits are: Data[6], Data[10], Data[8], Data[3], Data[7], Data[5], Data[9], Data[11]

The symbolic expression is:
(((((((~((~(D[2]) & ~(D[1])) & ~(D[4])) | D[6]) & (~((D[2] & ~(D[1])) & ~(D[4])) | D[10])) & (~((~(D[2]) & D[1]) & ~(D[4])) | D[8])) & (~((D[2] & D[1]) & ~(D[4])) | D[3])) & (~((~(D[2]) & ~(D[1])) & D[4]) | D[7])) & (~((D[2] & ~(D[1])) & D[4]) | D[5])) & (~((~(D[2]) & D[1]) & D[4]) | D[9])) & (~((D[2] & D[1]) & D[4]) | D[11])

*)

FUNCTION_BLOCK F_CollectInput
  VAR_IN_OUT
      Data : ARRAY[1..15] OF BOOL;
  END_VAR
  VAR_INPUT
      TICK  : BOOL := 0;
      IN1   : BOOL := 0;
      IN2   : BOOL := 0;
      IN3   : BOOL := 0;
      IN4   : BOOL := 0;
      IN5   : BOOL := 0;
      RESET : BOOL := FALSE;
  END_VAR
  VAR_OUTPUT
      Finished : BOOL;
  END_VAR
  VAR
      j    : USINT := 1;
      tock : BOOL  := 0;
  END_VAR
  IF NOT RESET AND tock = NOT TICK THEN
      Data[j]   := IN1;
      Data[j+1] := IN2;
      Data[j+2] := IN3;
      Data[j+3] := IN4;
      Data[j+4] := IN5;
      j := j + 5;
      tock := TICK;
  ELSE
      j := 1;
      tock := 0;
  END_IF;
  Finished := (j > 15);
END_FUNCTION_BLOCK

PROGRAM Boiler
  VAR
    Data  : ARRAY[1..15] OF BOOL;
    Ready : BOOL;
    CollectInput : F_CollectInput;
  END_VAR
  VAR
    TICK     AT %IX1.0 : BOOL;
    IN1      AT %IX0.3 : BOOL;
    IN2      AT %IX0.4 : BOOL;
    IN3      AT %IX0.5 : BOOL;
    IN4      AT %IX0.6 : BOOL;
    IN5      AT %IX0.7 : BOOL;
    OutReady AT %QX0.0 : BOOL := FALSE;
    FeedNext AT %QX0.1 : BOOL := FALSE;
    Out      AT %QX0.2 : BOOL;
  END_VAR
  CollectInput(TICK:=TICK, IN1:=IN1, IN2:=IN2, IN3:=IN3, IN4:=IN4, IN5:=IN5);
  Ready := CollectInput.Finished;
  FeedNext := 1;
  IF Ready THEN
    Out := (((((((((NOT (((NOT D[2]) AND (NOT D[1])) AND (NOT D[4]))) OR D[6]) AND ((NOT ((D[2] AND (NOT D[1])) AND (NOT D[4]))) OR D[10])) AND ((NOT (((NOT D[2]) AND D[1]) AND (NOT D[4]))) OR D[8])) AND ((NOT ((D[2] AND D[1]) AND (NOT D[4]))) OR D[3])) AND ((NOT (((NOT D[2]) AND (NOT D[1])) AND D[4])) OR D[7])) AND ((NOT ((D[2] AND (NOT D[1])) AND D[4])) OR D[5])) AND ((NOT (((NOT D[2]) AND D[1]) AND D[4])) OR D[9])) AND ((NOT ((D[2] AND D[1]) AND D[4])) OR D[11]));
    OutReady := 1;
    CollectInput(RESET:=TRUE);
  END_IF;
END_PROGRAM

CONFIGURATION Config0
  RESOURCE Res0 ON PLC
    TASK task0(INTERVAL := T#20ms,PRIORITY := 0);
    PROGRAM instance0 WITH task0 : Boiler;
  END_RESOURCE
END_CONFIGURATION

(* ---- 3-MUX_vapor-slays-token.st ---- *)
(*
This code implements a shuffled multiplexer with 3 control bits.
The control bits are: Data[3], Data[1], Data[2]
The input bits are: Data[5], Data[4], Data[6], Data[10], Data[11], Data[8], Data[9], Data[7]

The symbolic expression is:
(((((((~((~(D[3]) & ~(D[1])) & ~(D[2])) | D[5]) & (~((D[3] & ~(D[1])) & ~(D[2])) | D[4])) & (~((~(D[3]) & D[1]) & ~(D[2])) | D[6])) & (~((D[3] & D[1]) & ~(D[2])) | D[10])) & (~((~(D[3]) & ~(D[1])) & D[2]) | D[11])) & (~((D[3] & ~(D[1])) & D[2]) | D[8])) & (~((~(D[3]) & D[1]) & D[2]) | D[9])) & (~((D[3] & D[1]) & D[2]) | D[7])

*)

FUNCTION_BLOCK F_CollectInput
  VAR_IN_OUT
      Data : ARRAY[1..15] OF BOOL;
  END_VAR
  VAR_INPUT
      TICK  : BOOL := 0;
      IN1   : BOOL := 0;
      IN2   : BOOL := 0;
      IN3   : BOOL := 0;
      IN4   : BOOL := 0;
      IN5   : BOOL := 0;
      RESET : BOOL := FALSE;
  END_VAR
  VAR_OUTPUT
      Finished : BOOL;
  END_VAR
  VAR
      j    : USINT := 1;
      tock : BOOL  := 0;
  END_VAR
  IF NOT RESET AND tock = NOT TICK THEN
      Data[j]   := IN1;
      Data[j+1] := IN2;
      Data[j+2] := IN3;
      Data[j+3] := IN4;
      Data[j+4] := IN5;
      j := j + 5;
      tock := TICK;
  ELSE
      j := 1;
      tock := 0;
  END_IF;
  Finished := (j > 15);
END_FUNCTION_BLOCK

PROGRAM Boiler
  VAR
    Data  : ARRAY[1..15] OF BOOL;
    Ready : BOOL;
    CollectInput : F_CollectInput;
  END_VAR
  VAR
    TICK     AT %IX1.0 : BOOL;
    IN1      AT %IX0.3 : BOOL;
    IN2      AT %IX0.4 : BOOL;
    IN3      AT %IX0.5 : BOOL;
    IN4      AT %IX0.6 : BOOL;
    IN5      AT %IX0.7 : BOOL;
    OutReady AT %QX0.0 : BOOL := FALSE;
    FeedNext AT %QX0.1 : BOOL := FALSE;
    Out      AT %QX0.2 : BOOL;
  END_VAR
  CollectInput(TICK:=TICK, IN1:=IN1, IN2:=IN2, IN3:=IN3, IN4:=IN4, IN5:=IN5);
  Ready := CollectInput.Finished;
  FeedNext := 1;
  IF Ready THEN
    Out := (((((((((NOT (((NOT D[3]) AND (NOT D[1])) AND (NOT D[2]))) OR D[5]) AND ((NOT ((D[3] AND (NOT D[1])) AND (NOT D[2]))) OR D[4])) AND ((NOT (((NOT D[3]) AND D[1]) AND (NOT D[2]))) OR D[6])) AND ((NOT ((D[3] AND D[1]) AND (NOT D[2]))) OR D[10])) AND ((NOT (((NOT D[3]) AND (NOT D[1])) AND D[2])) OR D[11])) AND ((NOT ((D[3] AND (NOT D[1])) AND D[2])) OR D[8])) AND ((NOT (((NOT D[3]) AND D[1]) AND D[2])) OR D[9])) AND ((NOT ((D[3] AND D[1]) AND D[2])) OR D[7]));
    OutReady := 1;
    CollectInput(RESET:=TRUE);
  END_IF;
END_PROGRAM

CONFIGURATION Config0
  RESOURCE Res0 ON PLC
    TASK task0(INTERVAL := T#20ms,PRIORITY := 0);
    PROGRAM instance0 WITH task0 : Boiler;
  END_RESOURCE
END_CONFIGURATION

(* ---- 3-MUX_vests-hands-shrub.st ---- *)
(*
This code implements a shuffled multiplexer with 3 control bits.
The control bits are: Data[2], Data[5], Data[1]
The input bits are: Data[10], Data[6], Data[3], Data[4], Data[7], Data[9], Data[8], Data[11]

The symbolic expression is:
(((((((~((~(D[2]) & ~(D[5])) & ~(D[1])) | D[10]) & (~((D[2] & ~(D[5])) & ~(D[1])) | D[6])) & (~((~(D[2]) & D[5]) & ~(D[1])) | D[3])) & (~((D[2] & D[5]) & ~(D[1])) | D[4])) & (~((~(D[2]) & ~(D[5])) & D[1]) | D[7])) & (~((D[2] & ~(D[5])) & D[1]) | D[9])) & (~((~(D[2]) & D[5]) & D[1]) | D[8])) & (~((D[2] & D[5]) & D[1]) | D[11])

*)

FUNCTION_BLOCK F_CollectInput
  VAR_IN_OUT
      Data : ARRAY[1..15] OF BOOL;
  END_VAR
  VAR_INPUT
      TICK  : BOOL := 0;
      IN1   : BOOL := 0;
      IN2   : BOOL := 0;
      IN3   : BOOL := 0;
      IN4   : BOOL := 0;
      IN5   : BOOL := 0;
      RESET : BOOL := FALSE;
  END_VAR
  VAR_OUTPUT
      Finished : BOOL;
  END_VAR
  VAR
      j    : USINT := 1;
      tock : BOOL  := 0;
  END_VAR
  IF NOT RESET AND tock = NOT TICK THEN
      Data[j]   := IN1;
      Data[j+1] := IN2;
      Data[j+2] := IN3;
      Data[j+3] := IN4;
      Data[j+4] := IN5;
      j := j + 5;
      tock := TICK;
  ELSE
      j := 1;
      tock := 0;
  END_IF;
  Finished := (j > 15);
END_FUNCTION_BLOCK

PROGRAM Boiler
  VAR
    Data  : ARRAY[1..15] OF BOOL;
    Ready : BOOL;
    CollectInput : F_CollectInput;
  END_VAR
  VAR
    TICK     AT %IX1.0 : BOOL;
    IN1      AT %IX0.3 : BOOL;
    IN2      AT %IX0.4 : BOOL;
    IN3      AT %IX0.5 : BOOL;
    IN4      AT %IX0.6 : BOOL;
    IN5      AT %IX0.7 : BOOL;
    OutReady AT %QX0.0 : BOOL := FALSE;
    FeedNext AT %QX0.1 : BOOL := FALSE;
    Out      AT %QX0.2 : BOOL;
  END_VAR
  CollectInput(TICK:=TICK, IN1:=IN1, IN2:=IN2, IN3:=IN3, IN4:=IN4, IN5:=IN5);
  Ready := CollectInput.Finished;
  FeedNext := 1;
  IF Ready THEN
    Out := (((((((((NOT (((NOT D[2]) AND (NOT D[5])) AND (NOT D[1]))) OR D[10]) AND ((NOT ((D[2] AND (NOT D[5])) AND (NOT D[1]))) OR D[6])) AND ((NOT (((NOT D[2]) AND D[5]) AND (NOT D[1]))) OR D[3])) AND ((NOT ((D[2] AND D[5]) AND (NOT D[1]))) OR D[4])) AND ((NOT (((NOT D[2]) AND (NOT D[5])) AND D[1])) OR D[7])) AND ((NOT ((D[2] AND (NOT D[5])) AND D[1])) OR D[9])) AND ((NOT (((NOT D[2]) AND D[5]) AND D[1])) OR D[8])) AND ((NOT ((D[2] AND D[5]) AND D[1])) OR D[11]));
    OutReady := 1;
    CollectInput(RESET:=TRUE);
  END_IF;
END_PROGRAM

CONFIGURATION Config0
  RESOURCE Res0 ON PLC
    TASK task0(INTERVAL := T#20ms,PRIORITY := 0);
    PROGRAM instance0 WITH task0 : Boiler;
  END_RESOURCE
END_CONFIGURATION

(* ---- 3-MUX_viers-toons-sexed.st ---- *)
(*
This code implements a shuffled multiplexer with 3 control bits.
The control bits are: Data[1], Data[7], Data[3]
The input bits are: Data[2], Data[4], Data[5], Data[6], Data[8], Data[9], Data[11], Data[10]

The symbolic expression is:
(((((((~((~(D[1]) & ~(D[7])) & ~(D[3])) | D[2]) & (~((D[1] & ~(D[7])) & ~(D[3])) | D[4])) & (~((~(D[1]) & D[7]) & ~(D[3])) | D[5])) & (~((D[1] & D[7]) & ~(D[3])) | D[6])) & (~((~(D[1]) & ~(D[7])) & D[3]) | D[8])) & (~((D[1] & ~(D[7])) & D[3]) | D[9])) & (~((~(D[1]) & D[7]) & D[3]) | D[11])) & (~((D[1] & D[7]) & D[3]) | D[10])

*)

FUNCTION_BLOCK F_CollectInput
  VAR_IN_OUT
      Data : ARRAY[1..15] OF BOOL;
  END_VAR
  VAR_INPUT
      TICK  : BOOL := 0;
      IN1   : BOOL := 0;
      IN2   : BOOL := 0;
      IN3   : BOOL := 0;
      IN4   : BOOL := 0;
      IN5   : BOOL := 0;
      RESET : BOOL := FALSE;
  END_VAR
  VAR_OUTPUT
      Finished : BOOL;
  END_VAR
  VAR
      j    : USINT := 1;
      tock : BOOL  := 0;
  END_VAR
  IF NOT RESET AND tock = NOT TICK THEN
      Data[j]   := IN1;
      Data[j+1] := IN2;
      Data[j+2] := IN3;
      Data[j+3] := IN4;
      Data[j+4] := IN5;
      j := j + 5;
      tock := TICK;
  ELSE
      j := 1;
      tock := 0;
  END_IF;
  Finished := (j > 15);
END_FUNCTION_BLOCK

PROGRAM Boiler
  VAR
    Data  : ARRAY[1..15] OF BOOL;
    Ready : BOOL;
    CollectInput : F_CollectInput;
  END_VAR
  VAR
    TICK     AT %IX1.0 : BOOL;
    IN1      AT %IX0.3 : BOOL;
    IN2      AT %IX0.4 : BOOL;
    IN3      AT %IX0.5 : BOOL;
    IN4      AT %IX0.6 : BOOL;
    IN5      AT %IX0.7 : BOOL;
    OutReady AT %QX0.0 : BOOL := FALSE;
    FeedNext AT %QX0.1 : BOOL := FALSE;
    Out      AT %QX0.2 : BOOL;
  END_VAR
  CollectInput(TICK:=TICK, IN1:=IN1, IN2:=IN2, IN3:=IN3, IN4:=IN4, IN5:=IN5);
  Ready := CollectInput.Finished;
  FeedNext := 1;
  IF Ready THEN
    Out := (((((((((NOT (((NOT D[1]) AND (NOT D[7])) AND (NOT D[3]))) OR D[2]) AND ((NOT ((D[1] AND (NOT D[7])) AND (NOT D[3]))) OR D[4])) AND ((NOT (((NOT D[1]) AND D[7]) AND (NOT D[3]))) OR D[5])) AND ((NOT ((D[1] AND D[7]) AND (NOT D[3]))) OR D[6])) AND ((NOT (((NOT D[1]) AND (NOT D[7])) AND D[3])) OR D[8])) AND ((NOT ((D[1] AND (NOT D[7])) AND D[3])) OR D[9])) AND ((NOT (((NOT D[1]) AND D[7]) AND D[3])) OR D[11])) AND ((NOT ((D[1] AND D[7]) AND D[3])) OR D[10]));
    OutReady := 1;
    CollectInput(RESET:=TRUE);
  END_IF;
END_PROGRAM

CONFIGURATION Config0
  RESOURCE Res0 ON PLC
    TASK task0(INTERVAL := T#20ms,PRIORITY := 0);
    PROGRAM instance0 WITH task0 : Boiler;
  END_RESOURCE
END_CONFIGURATION

(* ---- 3-MUX_viral-hades-whips.st ---- *)
(*
This code implements a shuffled multiplexer with 3 control bits.
The control bits are: Data[3], Data[1], Data[2]
The input bits are: Data[6], Data[4], Data[5], Data[8], Data[7], Data[10], Data[9], Data[11]

The symbolic expression is:
(((((((~((~(D[3]) & ~(D[1])) & ~(D[2])) | D[6]) & (~((D[3] & ~(D[1])) & ~(D[2])) | D[4])) & (~((~(D[3]) & D[1]) & ~(D[2])) | D[5])) & (~((D[3] & D[1]) & ~(D[2])) | D[8])) & (~((~(D[3]) & ~(D[1])) & D[2]) | D[7])) & (~((D[3] & ~(D[1])) & D[2]) | D[10])) & (~((~(D[3]) & D[1]) & D[2]) | D[9])) & (~((D[3] & D[1]) & D[2]) | D[11])

*)

FUNCTION_BLOCK F_CollectInput
  VAR_IN_OUT
      Data : ARRAY[1..15] OF BOOL;
  END_VAR
  VAR_INPUT
      TICK  : BOOL := 0;
      IN1   : BOOL := 0;
      IN2   : BOOL := 0;
      IN3   : BOOL := 0;
      IN4   : BOOL := 0;
      IN5   : BOOL := 0;
      RESET : BOOL := FALSE;
  END_VAR
  VAR_OUTPUT
      Finished : BOOL;
  END_VAR
  VAR
      j    : USINT := 1;
      tock : BOOL  := 0;
  END_VAR
  IF NOT RESET AND tock = NOT TICK THEN
      Data[j]   := IN1;
      Data[j+1] := IN2;
      Data[j+2] := IN3;
      Data[j+3] := IN4;
      Data[j+4] := IN5;
      j := j + 5;
      tock := TICK;
  ELSE
      j := 1;
      tock := 0;
  END_IF;
  Finished := (j > 15);
END_FUNCTION_BLOCK

PROGRAM Boiler
  VAR
    Data  : ARRAY[1..15] OF BOOL;
    Ready : BOOL;
    CollectInput : F_CollectInput;
  END_VAR
  VAR
    TICK     AT %IX1.0 : BOOL;
    IN1      AT %IX0.3 : BOOL;
    IN2      AT %IX0.4 : BOOL;
    IN3      AT %IX0.5 : BOOL;
    IN4      AT %IX0.6 : BOOL;
    IN5      AT %IX0.7 : BOOL;
    OutReady AT %QX0.0 : BOOL := FALSE;
    FeedNext AT %QX0.1 : BOOL := FALSE;
    Out      AT %QX0.2 : BOOL;
  END_VAR
  CollectInput(TICK:=TICK, IN1:=IN1, IN2:=IN2, IN3:=IN3, IN4:=IN4, IN5:=IN5);
  Ready := CollectInput.Finished;
  FeedNext := 1;
  IF Ready THEN
    Out := (((((((((NOT (((NOT D[3]) AND (NOT D[1])) AND (NOT D[2]))) OR D[6]) AND ((NOT ((D[3] AND (NOT D[1])) AND (NOT D[2]))) OR D[4])) AND ((NOT (((NOT D[3]) AND D[1]) AND (NOT D[2]))) OR D[5])) AND ((NOT ((D[3] AND D[1]) AND (NOT D[2]))) OR D[8])) AND ((NOT (((NOT D[3]) AND (NOT D[1])) AND D[2])) OR D[7])) AND ((NOT ((D[3] AND (NOT D[1])) AND D[2])) OR D[10])) AND ((NOT (((NOT D[3]) AND D[1]) AND D[2])) OR D[9])) AND ((NOT ((D[3] AND D[1]) AND D[2])) OR D[11]));
    OutReady := 1;
    CollectInput(RESET:=TRUE);
  END_IF;
END_PROGRAM

CONFIGURATION Config0
  RESOURCE Res0 ON PLC
    TASK task0(INTERVAL := T#20ms,PRIORITY := 0);
    PROGRAM instance0 WITH task0 : Boiler;
  END_RESOURCE
END_CONFIGURATION

(* ---- 3-MUX_waltz-goers-witty.st ---- *)
(*
This code implements a shuffled multiplexer with 3 control bits.
The control bits are: Data[3], Data[1], Data[2]
The input bits are: Data[4], Data[6], Data[5], Data[7], Data[8], Data[9], Data[11], Data[10]

The symbolic expression is:
(((((((~((~(D[3]) & ~(D[1])) & ~(D[2])) | D[4]) & (~((D[3] & ~(D[1])) & ~(D[2])) | D[6])) & (~((~(D[3]) & D[1]) & ~(D[2])) | D[5])) & (~((D[3] & D[1]) & ~(D[2])) | D[7])) & (~((~(D[3]) & ~(D[1])) & D[2]) | D[8])) & (~((D[3] & ~(D[1])) & D[2]) | D[9])) & (~((~(D[3]) & D[1]) & D[2]) | D[11])) & (~((D[3] & D[1]) & D[2]) | D[10])

*)

FUNCTION_BLOCK F_CollectInput
  VAR_IN_OUT
      Data : ARRAY[1..15] OF BOOL;
  END_VAR
  VAR_INPUT
      TICK  : BOOL := 0;
      IN1   : BOOL := 0;
      IN2   : BOOL := 0;
      IN3   : BOOL := 0;
      IN4   : BOOL := 0;
      IN5   : BOOL := 0;
      RESET : BOOL := FALSE;
  END_VAR
  VAR_OUTPUT
      Finished : BOOL;
  END_VAR
  VAR
      j    : USINT := 1;
      tock : BOOL  := 0;
  END_VAR
  IF NOT RESET AND tock = NOT TICK THEN
      Data[j]   := IN1;
      Data[j+1] := IN2;
      Data[j+2] := IN3;
      Data[j+3] := IN4;
      Data[j+4] := IN5;
      j := j + 5;
      tock := TICK;
  ELSE
      j := 1;
      tock := 0;
  END_IF;
  Finished := (j > 15);
END_FUNCTION_BLOCK

PROGRAM Boiler
  VAR
    Data  : ARRAY[1..15] OF BOOL;
    Ready : BOOL;
    CollectInput : F_CollectInput;
  END_VAR
  VAR
    TICK     AT %IX1.0 : BOOL;
    IN1      AT %IX0.3 : BOOL;
    IN2      AT %IX0.4 : BOOL;
    IN3      AT %IX0.5 : BOOL;
    IN4      AT %IX0.6 : BOOL;
    IN5      AT %IX0.7 : BOOL;
    OutReady AT %QX0.0 : BOOL := FALSE;
    FeedNext AT %QX0.1 : BOOL := FALSE;
    Out      AT %QX0.2 : BOOL;
  END_VAR
  CollectInput(TICK:=TICK, IN1:=IN1, IN2:=IN2, IN3:=IN3, IN4:=IN4, IN5:=IN5);
  Ready := CollectInput.Finished;
  FeedNext := 1;
  IF Ready THEN
    Out := (((((((((NOT (((NOT D[3]) AND (NOT D[1])) AND (NOT D[2]))) OR D[4]) AND ((NOT ((D[3] AND (NOT D[1])) AND (NOT D[2]))) OR D[6])) AND ((NOT (((NOT D[3]) AND D[1]) AND (NOT D[2]))) OR D[5])) AND ((NOT ((D[3] AND D[1]) AND (NOT D[2]))) OR D[7])) AND ((NOT (((NOT D[3]) AND (NOT D[1])) AND D[2])) OR D[8])) AND ((NOT ((D[3] AND (NOT D[1])) AND D[2])) OR D[9])) AND ((NOT (((NOT D[3]) AND D[1]) AND D[2])) OR D[11])) AND ((NOT ((D[3] AND D[1]) AND D[2])) OR D[10]));
    OutReady := 1;
    CollectInput(RESET:=TRUE);
  END_IF;
END_PROGRAM

CONFIGURATION Config0
  RESOURCE Res0 ON PLC
    TASK task0(INTERVAL := T#20ms,PRIORITY := 0);
    PROGRAM instance0 WITH task0 : Boiler;
  END_RESOURCE
END_CONFIGURATION

(* ---- 3-MUX_wards-sidle-paged.st ---- *)
(*
This code implements a shuffled multiplexer with 3 control bits.
The control bits are: Data[1], Data[2], Data[3]
The input bits are: Data[4], Data[8], Data[6], Data[7], Data[9], Data[5], Data[10], Data[11]

The symbolic expression is:
(((((((~((~(D[1]) & ~(D[2])) & ~(D[3])) | D[4]) & (~((D[1] & ~(D[2])) & ~(D[3])) | D[8])) & (~((~(D[1]) & D[2]) & ~(D[3])) | D[6])) & (~((D[1] & D[2]) & ~(D[3])) | D[7])) & (~((~(D[1]) & ~(D[2])) & D[3]) | D[9])) & (~((D[1] & ~(D[2])) & D[3]) | D[5])) & (~((~(D[1]) & D[2]) & D[3]) | D[10])) & (~((D[1] & D[2]) & D[3]) | D[11])

*)

FUNCTION_BLOCK F_CollectInput
  VAR_IN_OUT
      Data : ARRAY[1..15] OF BOOL;
  END_VAR
  VAR_INPUT
      TICK  : BOOL := 0;
      IN1   : BOOL := 0;
      IN2   : BOOL := 0;
      IN3   : BOOL := 0;
      IN4   : BOOL := 0;
      IN5   : BOOL := 0;
      RESET : BOOL := FALSE;
  END_VAR
  VAR_OUTPUT
      Finished : BOOL;
  END_VAR
  VAR
      j    : USINT := 1;
      tock : BOOL  := 0;
  END_VAR
  IF NOT RESET AND tock = NOT TICK THEN
      Data[j]   := IN1;
      Data[j+1] := IN2;
      Data[j+2] := IN3;
      Data[j+3] := IN4;
      Data[j+4] := IN5;
      j := j + 5;
      tock := TICK;
  ELSE
      j := 1;
      tock := 0;
  END_IF;
  Finished := (j > 15);
END_FUNCTION_BLOCK

PROGRAM Boiler
  VAR
    Data  : ARRAY[1..15] OF BOOL;
    Ready : BOOL;
    CollectInput : F_CollectInput;
  END_VAR
  VAR
    TICK     AT %IX1.0 : BOOL;
    IN1      AT %IX0.3 : BOOL;
    IN2      AT %IX0.4 : BOOL;
    IN3      AT %IX0.5 : BOOL;
    IN4      AT %IX0.6 : BOOL;
    IN5      AT %IX0.7 : BOOL;
    OutReady AT %QX0.0 : BOOL := FALSE;
    FeedNext AT %QX0.1 : BOOL := FALSE;
    Out      AT %QX0.2 : BOOL;
  END_VAR
  CollectInput(TICK:=TICK, IN1:=IN1, IN2:=IN2, IN3:=IN3, IN4:=IN4, IN5:=IN5);
  Ready := CollectInput.Finished;
  FeedNext := 1;
  IF Ready THEN
    Out := (((((((((NOT (((NOT D[1]) AND (NOT D[2])) AND (NOT D[3]))) OR D[4]) AND ((NOT ((D[1] AND (NOT D[2])) AND (NOT D[3]))) OR D[8])) AND ((NOT (((NOT D[1]) AND D[2]) AND (NOT D[3]))) OR D[6])) AND ((NOT ((D[1] AND D[2]) AND (NOT D[3]))) OR D[7])) AND ((NOT (((NOT D[1]) AND (NOT D[2])) AND D[3])) OR D[9])) AND ((NOT ((D[1] AND (NOT D[2])) AND D[3])) OR D[5])) AND ((NOT (((NOT D[1]) AND D[2]) AND D[3])) OR D[10])) AND ((NOT ((D[1] AND D[2]) AND D[3])) OR D[11]));
    OutReady := 1;
    CollectInput(RESET:=TRUE);
  END_IF;
END_PROGRAM

CONFIGURATION Config0
  RESOURCE Res0 ON PLC
    TASK task0(INTERVAL := T#20ms,PRIORITY := 0);
    PROGRAM instance0 WITH task0 : Boiler;
  END_RESOURCE
END_CONFIGURATION

(* ---- 3-MUX_wefts-raise-fovea.st ---- *)
(*
This code implements a shuffled multiplexer with 3 control bits.
The control bits are: Data[1], Data[3], Data[2]
The input bits are: Data[6], Data[4], Data[5], Data[7], Data[10], Data[8], Data[9], Data[11]

The symbolic expression is:
(((((((~((~(D[1]) & ~(D[3])) & ~(D[2])) | D[6]) & (~((D[1] & ~(D[3])) & ~(D[2])) | D[4])) & (~((~(D[1]) & D[3]) & ~(D[2])) | D[5])) & (~((D[1] & D[3]) & ~(D[2])) | D[7])) & (~((~(D[1]) & ~(D[3])) & D[2]) | D[10])) & (~((D[1] & ~(D[3])) & D[2]) | D[8])) & (~((~(D[1]) & D[3]) & D[2]) | D[9])) & (~((D[1] & D[3]) & D[2]) | D[11])

*)

FUNCTION_BLOCK F_CollectInput
  VAR_IN_OUT
      Data : ARRAY[1..15] OF BOOL;
  END_VAR
  VAR_INPUT
      TICK  : BOOL := 0;
      IN1   : BOOL := 0;
      IN2   : BOOL := 0;
      IN3   : BOOL := 0;
      IN4   : BOOL := 0;
      IN5   : BOOL := 0;
      RESET : BOOL := FALSE;
  END_VAR
  VAR_OUTPUT
      Finished : BOOL;
  END_VAR
  VAR
      j    : USINT := 1;
      tock : BOOL  := 0;
  END_VAR
  IF NOT RESET AND tock = NOT TICK THEN
      Data[j]   := IN1;
      Data[j+1] := IN2;
      Data[j+2] := IN3;
      Data[j+3] := IN4;
      Data[j+4] := IN5;
      j := j + 5;
      tock := TICK;
  ELSE
      j := 1;
      tock := 0;
  END_IF;
  Finished := (j > 15);
END_FUNCTION_BLOCK

PROGRAM Boiler
  VAR
    Data  : ARRAY[1..15] OF BOOL;
    Ready : BOOL;
    CollectInput : F_CollectInput;
  END_VAR
  VAR
    TICK     AT %IX1.0 : BOOL;
    IN1      AT %IX0.3 : BOOL;
    IN2      AT %IX0.4 : BOOL;
    IN3      AT %IX0.5 : BOOL;
    IN4      AT %IX0.6 : BOOL;
    IN5      AT %IX0.7 : BOOL;
    OutReady AT %QX0.0 : BOOL := FALSE;
    FeedNext AT %QX0.1 : BOOL := FALSE;
    Out      AT %QX0.2 : BOOL;
  END_VAR
  CollectInput(TICK:=TICK, IN1:=IN1, IN2:=IN2, IN3:=IN3, IN4:=IN4, IN5:=IN5);
  Ready := CollectInput.Finished;
  FeedNext := 1;
  IF Ready THEN
    Out := (((((((((NOT (((NOT D[1]) AND (NOT D[3])) AND (NOT D[2]))) OR D[6]) AND ((NOT ((D[1] AND (NOT D[3])) AND (NOT D[2]))) OR D[4])) AND ((NOT (((NOT D[1]) AND D[3]) AND (NOT D[2]))) OR D[5])) AND ((NOT ((D[1] AND D[3]) AND (NOT D[2]))) OR D[7])) AND ((NOT (((NOT D[1]) AND (NOT D[3])) AND D[2])) OR D[10])) AND ((NOT ((D[1] AND (NOT D[3])) AND D[2])) OR D[8])) AND ((NOT (((NOT D[1]) AND D[3]) AND D[2])) OR D[9])) AND ((NOT ((D[1] AND D[3]) AND D[2])) OR D[11]));
    OutReady := 1;
    CollectInput(RESET:=TRUE);
  END_IF;
END_PROGRAM

CONFIGURATION Config0
  RESOURCE Res0 ON PLC
    TASK task0(INTERVAL := T#20ms,PRIORITY := 0);
    PROGRAM instance0 WITH task0 : Boiler;
  END_RESOURCE
END_CONFIGURATION

(* ---- 3-MUX_whelm-blink-visit.st ---- *)
(*
This code implements a shuffled multiplexer with 3 control bits.
The control bits are: Data[2], Data[1], Data[3]
The input bits are: Data[4], Data[5], Data[8], Data[6], Data[10], Data[7], Data[9], Data[11]

The symbolic expression is:
(((((((~((~(D[2]) & ~(D[1])) & ~(D[3])) | D[4]) & (~((D[2] & ~(D[1])) & ~(D[3])) | D[5])) & (~((~(D[2]) & D[1]) & ~(D[3])) | D[8])) & (~((D[2] & D[1]) & ~(D[3])) | D[6])) & (~((~(D[2]) & ~(D[1])) & D[3]) | D[10])) & (~((D[2] & ~(D[1])) & D[3]) | D[7])) & (~((~(D[2]) & D[1]) & D[3]) | D[9])) & (~((D[2] & D[1]) & D[3]) | D[11])

*)

FUNCTION_BLOCK F_CollectInput
  VAR_IN_OUT
      Data : ARRAY[1..15] OF BOOL;
  END_VAR
  VAR_INPUT
      TICK  : BOOL := 0;
      IN1   : BOOL := 0;
      IN2   : BOOL := 0;
      IN3   : BOOL := 0;
      IN4   : BOOL := 0;
      IN5   : BOOL := 0;
      RESET : BOOL := FALSE;
  END_VAR
  VAR_OUTPUT
      Finished : BOOL;
  END_VAR
  VAR
      j    : USINT := 1;
      tock : BOOL  := 0;
  END_VAR
  IF NOT RESET AND tock = NOT TICK THEN
      Data[j]   := IN1;
      Data[j+1] := IN2;
      Data[j+2] := IN3;
      Data[j+3] := IN4;
      Data[j+4] := IN5;
      j := j + 5;
      tock := TICK;
  ELSE
      j := 1;
      tock := 0;
  END_IF;
  Finished := (j > 15);
END_FUNCTION_BLOCK

PROGRAM Boiler
  VAR
    Data  : ARRAY[1..15] OF BOOL;
    Ready : BOOL;
    CollectInput : F_CollectInput;
  END_VAR
  VAR
    TICK     AT %IX1.0 : BOOL;
    IN1      AT %IX0.3 : BOOL;
    IN2      AT %IX0.4 : BOOL;
    IN3      AT %IX0.5 : BOOL;
    IN4      AT %IX0.6 : BOOL;
    IN5      AT %IX0.7 : BOOL;
    OutReady AT %QX0.0 : BOOL := FALSE;
    FeedNext AT %QX0.1 : BOOL := FALSE;
    Out      AT %QX0.2 : BOOL;
  END_VAR
  CollectInput(TICK:=TICK, IN1:=IN1, IN2:=IN2, IN3:=IN3, IN4:=IN4, IN5:=IN5);
  Ready := CollectInput.Finished;
  FeedNext := 1;
  IF Ready THEN
    Out := (((((((((NOT (((NOT D[2]) AND (NOT D[1])) AND (NOT D[3]))) OR D[4]) AND ((NOT ((D[2] AND (NOT D[1])) AND (NOT D[3]))) OR D[5])) AND ((NOT (((NOT D[2]) AND D[1]) AND (NOT D[3]))) OR D[8])) AND ((NOT ((D[2] AND D[1]) AND (NOT D[3]))) OR D[6])) AND ((NOT (((NOT D[2]) AND (NOT D[1])) AND D[3])) OR D[10])) AND ((NOT ((D[2] AND (NOT D[1])) AND D[3])) OR D[7])) AND ((NOT (((NOT D[2]) AND D[1]) AND D[3])) OR D[9])) AND ((NOT ((D[2] AND D[1]) AND D[3])) OR D[11]));
    OutReady := 1;
    CollectInput(RESET:=TRUE);
  END_IF;
END_PROGRAM

CONFIGURATION Config0
  RESOURCE Res0 ON PLC
    TASK task0(INTERVAL := T#20ms,PRIORITY := 0);
    PROGRAM instance0 WITH task0 : Boiler;
  END_RESOURCE
END_CONFIGURATION

(* ---- 3-MUX_woods-fores-femme.st ---- *)
(*
This code implements a shuffled multiplexer with 3 control bits.
The control bits are: Data[3], Data[2], Data[1]
The input bits are: Data[6], Data[7], Data[8], Data[9], Data[10], Data[11], Data[4], Data[5]

The symbolic expression is:
(((((((~((~(D[3]) & ~(D[2])) & ~(D[1])) | D[6]) & (~((D[3] & ~(D[2])) & ~(D[1])) | D[7])) & (~((~(D[3]) & D[2]) & ~(D[1])) | D[8])) & (~((D[3] & D[2]) & ~(D[1])) | D[9])) & (~((~(D[3]) & ~(D[2])) & D[1]) | D[10])) & (~((D[3] & ~(D[2])) & D[1]) | D[11])) & (~((~(D[3]) & D[2]) & D[1]) | D[4])) & (~((D[3] & D[2]) & D[1]) | D[5])

*)

FUNCTION_BLOCK F_CollectInput
  VAR_IN_OUT
      Data : ARRAY[1..15] OF BOOL;
  END_VAR
  VAR_INPUT
      TICK  : BOOL := 0;
      IN1   : BOOL := 0;
      IN2   : BOOL := 0;
      IN3   : BOOL := 0;
      IN4   : BOOL := 0;
      IN5   : BOOL := 0;
      RESET : BOOL := FALSE;
  END_VAR
  VAR_OUTPUT
      Finished : BOOL;
  END_VAR
  VAR
      j    : USINT := 1;
      tock : BOOL  := 0;
  END_VAR
  IF NOT RESET AND tock = NOT TICK THEN
      Data[j]   := IN1;
      Data[j+1] := IN2;
      Data[j+2] := IN3;
      Data[j+3] := IN4;
      Data[j+4] := IN5;
      j := j + 5;
      tock := TICK;
  ELSE
      j := 1;
      tock := 0;
  END_IF;
  Finished := (j > 15);
END_FUNCTION_BLOCK

PROGRAM Boiler
  VAR
    Data  : ARRAY[1..15] OF BOOL;
    Ready : BOOL;
    CollectInput : F_CollectInput;
  END_VAR
  VAR
    TICK     AT %IX1.0 : BOOL;
    IN1      AT %IX0.3 : BOOL;
    IN2      AT %IX0.4 : BOOL;
    IN3      AT %IX0.5 : BOOL;
    IN4      AT %IX0.6 : BOOL;
    IN5      AT %IX0.7 : BOOL;
    OutReady AT %QX0.0 : BOOL := FALSE;
    FeedNext AT %QX0.1 : BOOL := FALSE;
    Out      AT %QX0.2 : BOOL;
  END_VAR
  CollectInput(TICK:=TICK, IN1:=IN1, IN2:=IN2, IN3:=IN3, IN4:=IN4, IN5:=IN5);
  Ready := CollectInput.Finished;
  FeedNext := 1;
  IF Ready THEN
    Out := (((((((((NOT (((NOT D[3]) AND (NOT D[2])) AND (NOT D[1]))) OR D[6]) AND ((NOT ((D[3] AND (NOT D[2])) AND (NOT D[1]))) OR D[7])) AND ((NOT (((NOT D[3]) AND D[2]) AND (NOT D[1]))) OR D[8])) AND ((NOT ((D[3] AND D[2]) AND (NOT D[1]))) OR D[9])) AND ((NOT (((NOT D[3]) AND (NOT D[2])) AND D[1])) OR D[10])) AND ((NOT ((D[3] AND (NOT D[2])) AND D[1])) OR D[11])) AND ((NOT (((NOT D[3]) AND D[2]) AND D[1])) OR D[4])) AND ((NOT ((D[3] AND D[2]) AND D[1])) OR D[5]));
    OutReady := 1;
    CollectInput(RESET:=TRUE);
  END_IF;
END_PROGRAM

CONFIGURATION Config0
  RESOURCE Res0 ON PLC
    TASK task0(INTERVAL := T#20ms,PRIORITY := 0);
    PROGRAM instance0 WITH task0 : Boiler;
  END_RESOURCE
END_CONFIGURATION

(* ---- 3-MUX_zeros-regal-ocher.st ---- *)
(*
This code implements a shuffled multiplexer with 3 control bits.
The control bits are: Data[1], Data[2], Data[5]
The input bits are: Data[3], Data[7], Data[4], Data[8], Data[9], Data[6], Data[11], Data[10]

The symbolic expression is:
(((((((~((~(D[1]) & ~(D[2])) & ~(D[5])) | D[3]) & (~((D[1] & ~(D[2])) & ~(D[5])) | D[7])) & (~((~(D[1]) & D[2]) & ~(D[5])) | D[4])) & (~((D[1] & D[2]) & ~(D[5])) | D[8])) & (~((~(D[1]) & ~(D[2])) & D[5]) | D[9])) & (~((D[1] & ~(D[2])) & D[5]) | D[6])) & (~((~(D[1]) & D[2]) & D[5]) | D[11])) & (~((D[1] & D[2]) & D[5]) | D[10])

*)

FUNCTION_BLOCK F_CollectInput
  VAR_IN_OUT
      Data : ARRAY[1..15] OF BOOL;
  END_VAR
  VAR_INPUT
      TICK  : BOOL := 0;
      IN1   : BOOL := 0;
      IN2   : BOOL := 0;
      IN3   : BOOL := 0;
      IN4   : BOOL := 0;
      IN5   : BOOL := 0;
      RESET : BOOL := FALSE;
  END_VAR
  VAR_OUTPUT
      Finished : BOOL;
  END_VAR
  VAR
      j    : USINT := 1;
      tock : BOOL  := 0;
  END_VAR
  IF NOT RESET AND tock = NOT TICK THEN
      Data[j]   := IN1;
      Data[j+1] := IN2;
      Data[j+2] := IN3;
      Data[j+3] := IN4;
      Data[j+4] := IN5;
      j := j + 5;
      tock := TICK;
  ELSE
      j := 1;
      tock := 0;
  END_IF;
  Finished := (j > 15);
END_FUNCTION_BLOCK

PROGRAM Boiler
  VAR
    Data  : ARRAY[1..15] OF BOOL;
    Ready : BOOL;
    CollectInput : F_CollectInput;
  END_VAR
  VAR
    TICK     AT %IX1.0 : BOOL;
    IN1      AT %IX0.3 : BOOL;
    IN2      AT %IX0.4 : BOOL;
    IN3      AT %IX0.5 : BOOL;
    IN4      AT %IX0.6 : BOOL;
    IN5      AT %IX0.7 : BOOL;
    OutReady AT %QX0.0 : BOOL := FALSE;
    FeedNext AT %QX0.1 : BOOL := FALSE;
    Out      AT %QX0.2 : BOOL;
  END_VAR
  CollectInput(TICK:=TICK, IN1:=IN1, IN2:=IN2, IN3:=IN3, IN4:=IN4, IN5:=IN5);
  Ready := CollectInput.Finished;
  FeedNext := 1;
  IF Ready THEN
    Out := (((((((((NOT (((NOT D[1]) AND (NOT D[2])) AND (NOT D[5]))) OR D[3]) AND ((NOT ((D[1] AND (NOT D[2])) AND (NOT D[5]))) OR D[7])) AND ((NOT (((NOT D[1]) AND D[2]) AND (NOT D[5]))) OR D[4])) AND ((NOT ((D[1] AND D[2]) AND (NOT D[5]))) OR D[8])) AND ((NOT (((NOT D[1]) AND (NOT D[2])) AND D[5])) OR D[9])) AND ((NOT ((D[1] AND (NOT D[2])) AND D[5])) OR D[6])) AND ((NOT (((NOT D[1]) AND D[2]) AND D[5])) OR D[11])) AND ((NOT ((D[1] AND D[2]) AND D[5])) OR D[10]));
    OutReady := 1;
    CollectInput(RESET:=TRUE);
  END_IF;
END_PROGRAM

CONFIGURATION Config0
  RESOURCE Res0 ON PLC
    TASK task0(INTERVAL := T#20ms,PRIORITY := 0);
    PROGRAM instance0 WITH task0 : Boiler;
  END_RESOURCE
END_CONFIGURATION
